// TIA Portal V20 export
FUNCTION_BLOCK "PR_TT-1MasterSeq_Soft2.0_workflow_b380e4"   // FB53, LAD
{ S7_Optimized_Access := 'TRUE' }
// stored: MemoryReserve 100, SetENOAutomatically false
   VAR_INPUT
      iAllStationProcessOver : Bool;
      iAutoRunning : Bool;
      iHiPotTestOver_1 : Bool;
      iHiPotTestOver_2 : Bool;
      iHiPot_RTR_1 : Bool;
      iHiPot_RTR_2 : Bool;
      iIndexOver : Bool;
      iIndex_RTR_Place1 : Bool;
      iIndex_RTR_Place2 : Bool;
      iOTS_Frm_Shuttle_1 : Bool;
      iOTS_Frm_Shuttle_2 : Bool;
      iOTS_Frm_TransferGantry : Bool;
      iOperatorAck : Bool;
      iPartPickOver : Bool;
      iPartPickOver_1 : Bool;
      iPartPickOver_2 : Bool;
      iPartPlaceByTransferGantry : Bool;
      iPartPlaceOver_IFGantry : Bool;
      iPartPlaceOver_IndexPlace1 : Bool;
      iPartPlaceOver_IndexPlace2 : Bool;
      iPartPresent_IFGantry : Bool;
      iPartPresent_Shuttle_1 : Bool;
      iPartPresent_Shuttle_2 : Bool;
      iPartPresent_TxGantry_1 : Bool;
      iPartPresent_TxGantry_2 : Bool;
      iRTR_Frm_TransferGantry_1 : Bool;
      iRTR_Frm_TransferGantry_2 : Bool;
      iReset_fault : Bool;
      iShuttleReadyToReceive : Bool;
      iSstMode : Bool;
      iSstPB : Bool;
   END_VAR
   VAR_OUTPUT
      qError : Array[1..1] of Bool;
      qInfeedGantry_PickStart : Bool;
      qInfeedGantry_PlaceStart : Bool;
      qShuttle_1PickStart : Bool;
      qShuttle_1PlaceStart : Bool;
      qShuttle_2PickStart : Bool;
      qShuttle_2PlaceStart : Bool;
      qTransferGantry1_PickStart : Bool;
      qTransferGantry1_PlaceStart : Bool;
      qTransferGantry2_PickStart : Bool;
      qTransferGantry2_PlaceStart : Bool;
   END_VAR
   VAR
      c10_ChkPartStsAtSubStn_T1 : Bool;
      c10_ChkPartStsAtSubStn_T2 : Bool;
      c10_ChkPartStsAtSubStn_T3 : Bool;
      c10_ChkPartStsAtSubStn_T4 : Bool;
      c10_ChkPartStsAtSubStn_T5 : Bool;
      c10_ChkPartStsAtSubStn_T6 : Bool;
      c10_ChkPartStsAtSubStn_T7 : Bool;
      c130_ChkPartPrsntStsShuttle2_T1 : Bool;
      c130_ChkPartPrsntStsShuttle2_T2 : Bool;
      c200_ChkPartPrsntTxGantry1_T1 : Bool;
      c200_ChkPartPrsntTxGantry1_T2 : Bool;
      c250_ChkPartPrsntTxGantry2_T1 : Bool;
      c250_ChkPartPrsntTxGantry2_T2 : Bool;
      c300_ChkPartPrsntIndexer_T1 : Bool;
      c300_ChkPartPrsntIndexer_T2 : Bool;
      c30_ChkPartStsIFGantry_T1 : Bool;
      c30_ChkPartStsIFGantry_T2 : Bool;
      c70_ChkPartPrsntStsShuttle1_T1 : Bool;
      c70_ChkPartPrsntStsShuttle1_T2 : Bool;
      StateNo : Int;
      s100_WtHiPotTestOver1 : Bool;
      s100_WtHiPotTestOver1_T1 : Bool;
      s10_ChkPartStsAtSubStn : Bool;
      s10_ChkPartStsAtSubStn_T1 : Bool;
      s10_ChkPartStsAtSubStn_T2 : Bool;
      s10_ChkPartStsAtSubStn_T3 : Bool;
      s10_ChkPartStsAtSubStn_T4 : Bool;
      s10_ChkPartStsAtSubStn_T5 : Bool;
      s10_ChkPartStsAtSubStn_T6 : Bool;
      s10_ChkPartStsAtSubStn_T7 : Bool;
      s110_WtTxGantryRTR1 : Bool;
      s110_WtTxGantryRTR1_T1 : Bool;
      s120_WtPartUnldOvrTxGantry1 : Bool;
      s120_WtPartUnldOvrTxGantry1_T1 : Bool;
      s130_ChkPartPrsntStsShuttle2 : Bool;
      s130_ChkPartPrsntStsShuttle2_T1 : Bool;
      s130_ChkPartPrsntStsShuttle2_T2 : Bool;
      s140_WtIFGantryPlacePart2 : Bool;
      s140_WtIFGantryPlacePart2_T1 : Bool;
      s150_WtHiPotRdyRcvPart2 : Bool;
      s150_WtHiPotRdyRcvPart2_T1 : Bool;
      s160_WtHiPotTestOver2 : Bool;
      s160_WtHiPotTestOver2_T1 : Bool;
      s170_WtTxGantryRTR2 : Bool;
      s170_WtTxGantryRTR2_T1 : Bool;
      s190_WtPartUnldOvrTxGantry2 : Bool;
      s190_WtPartUnldOvrTxGantry2_T1 : Bool;
      s1_WtResetRel : Bool;
      s1_WtResetRel_T1 : Bool;
      s200_ChkPartPrsntTxGantry1 : Bool;
      s200_ChkPartPrsntTxGantry1_T1 : Bool;
      s200_ChkPartPrsntTxGantry1_T2 : Bool;
      s20_WtOperatorAck : Bool;
      s20_WtOperatorAck_T1 : Bool;
      s210_WtShuttle1RdySendPal : Bool;
      s210_WtShuttle1RdySendPal_T1 : Bool;
      s220_WtPartPickTxGantry1 : Bool;
      s220_WtPartPickTxGantry1_T1 : Bool;
      s230_WtIndexRTRPlace1 : Bool;
      s230_WtIndexRTRPlace1_T1 : Bool;
      s240_WtPartPlaceOverIndexPlace1 : Bool;
      s240_WtPartPlaceOverIndexPlace1_T1 : Bool;
      s250_ChkPartPrsntTxGantry2 : Bool;
      s250_ChkPartPrsntTxGantry2_T1 : Bool;
      s250_ChkPartPrsntTxGantry2_T2 : Bool;
      s260_WtShuttle2RdySendPal : Bool;
      s260_WtShuttle2RdySendPal_T1 : Bool;
      s270_WtPartPickTxGantry2 : Bool;
      s270_WtPartPickTxGantry2_T1 : Bool;
      s280_WtIndexRTRPlace2 : Bool;
      s280_WtIndexRTRPlace2_T1 : Bool;
      s290_WtPartPlaceOverIndexPlace2 : Bool;
      s290_WtPartPlaceOverIndexPlace2_T1 : Bool;
      s300_ChkPartPrsntIndexer : Bool;
      s300_ChkPartPrsntIndexer_T1 : Bool;
      s300_ChkPartPrsntIndexer_T2 : Bool;
      s30_ChkPartStsIFGantry : Bool;
      s30_ChkPartStsIFGantry_T1 : Bool;
      s30_ChkPartStsIFGantry_T2 : Bool;
      s310_WtOTSFrmTxGantry : Bool;
      s310_WtOTSFrmTxGantry_T1 : Bool;
      s320_WtPartPlaceByTxGantry : Bool;
      s320_WtPartPlaceByTxGantry_T1 : Bool;
      s330_WtAllStnProcessOver : Bool;
      s330_WtAllStnProcessOver_T1 : Bool;
      s340_WtIndexOver : Bool;
      s340_WtIndexOver_T1 : Bool;
      s40_WtPartPickOverIFGantry : Bool;
      s40_WtPartPickOverIFGantry_T1 : Bool;
      s50_WtShuttleRdyRcvPart : Bool;
      s50_WtShuttleRdyRcvPart_T1 : Bool;
      s60_WtPartPlaceByGantry : Bool;
      s60_WtPartPlaceByGantry_T1 : Bool;
      s70_ChkPartPrsntStsShuttle1 : Bool;
      s70_ChkPartPrsntStsShuttle1_T1 : Bool;
      s70_ChkPartPrsntStsShuttle1_T2 : Bool;
      s80_WtIFGantryPlacePart : Bool;
      s80_WtIFGantryPlacePart_T1 : Bool;
      s90_WtHiPotRdyRcvPart1 : Bool;
      s90_WtHiPotRdyRcvPart1_T1 : Bool;
      sAbnormalCondition : Bool;
      sIndexerSeq : Bool;
      sInfeedGantry : Bool;
      sPartAbsentAtAllStn : Bool;
      sPartPrsntAtStn : Bool;
      sShuttle_1Seq : Bool;
      sShuttle_2Seq : Bool;
      sSst : Bool;
      sSstPulse : Bool;
      sSstRise : Bool;
      sStWtResetRel : Bool;
      sStWtResetRel_T1 : Bool;
      sTransferGantry_1Seq : Bool;
      sTransferGantry_2Seq : Bool;
   END_VAR
   VAR_TEMP
      tOne : Bool;
   END_VAR
   VAR_TEMP   // added for the SCL form of the ladder/FBD networks
      _w1 : Bool;
      _w2 : Bool;
      _w3 : Bool;
      _w4 : Bool;
      _w5 : Bool;
      _w6 : Bool;
   END_VAR
BEGIN

REGION Network 1
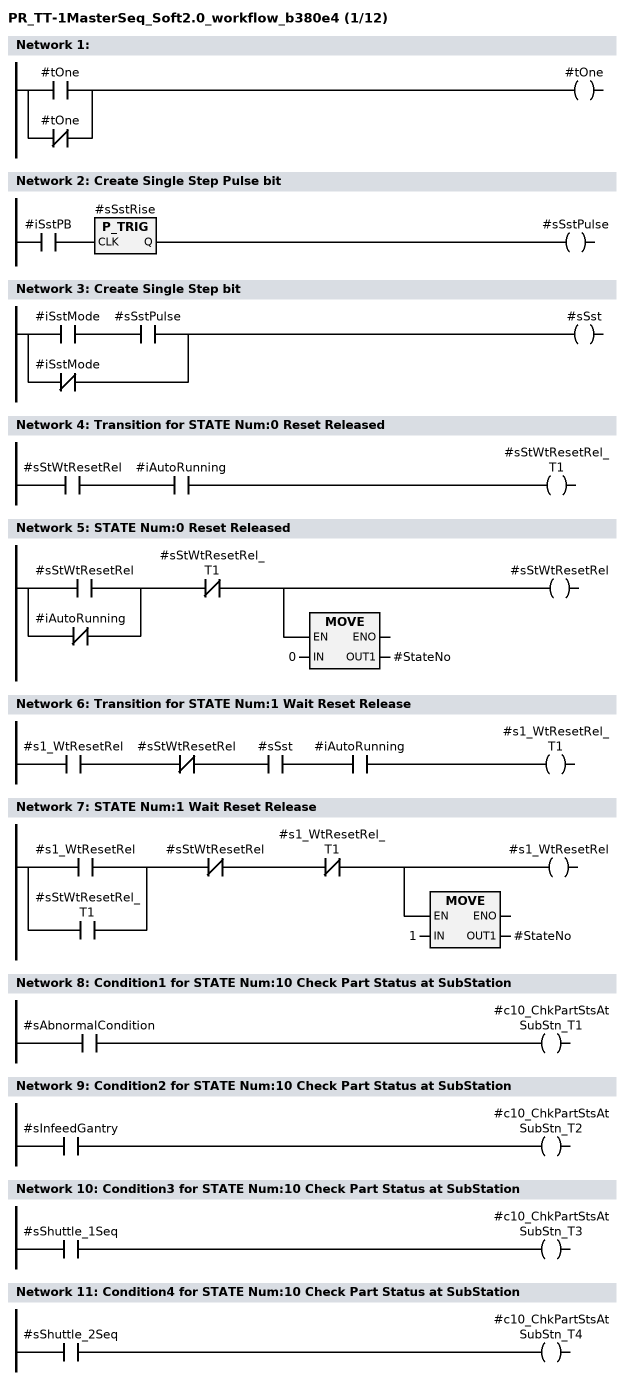
   RUNG wire#powerrail
      Contact( #tOne )
      wire#w1
      Coil( #tOne )
   END_RUNG
   RUNG wire#powerrail
      I_Contact( #tOne )
   END_RUNG wire#w1
   // the same network as SCL:
   #tOne := #tOne OR NOT #tOne;
END_REGION

REGION Network 2: Create Single Step Pulse bit
   RUNG wire#powerrail
      Contact( #iSstPB )
      P_Trig( #sSstRise )
      Coil( #sSstPulse )
   END_RUNG
   // the same network as SCL:
   #_w1 := #iSstPB AND NOT #sSstRise;   // rising edge
   #sSstRise := #iSstPB;
   #sSstPulse := #_w1;
END_REGION

REGION Network 3: Create Single Step bit
   RUNG wire#powerrail
      Contact( #iSstMode )
      Contact( #sSstPulse )
      wire#w1
      Coil( #sSst )
   END_RUNG
   RUNG wire#powerrail
      I_Contact( #iSstMode )
   END_RUNG wire#w1
   // the same network as SCL:
   #sSst := (#iSstMode AND #sSstPulse) OR NOT #iSstMode;
END_REGION

REGION Network 4: Transition for STATE Num:0 Reset Released
   RUNG wire#powerrail
      Contact( #sStWtResetRel )
      Contact( #iAutoRunning )
      Coil( #sStWtResetRel_T1 )
   END_RUNG
   // the same network as SCL:
   #sStWtResetRel_T1 := #sStWtResetRel AND #iAutoRunning;
END_REGION

REGION Network 5: STATE Num:0 Reset Released
   RUNG wire#powerrail
      Contact( #sStWtResetRel )
      wire#w1
      I_Contact( #sStWtResetRel_T1 )
      wire#w2
      Coil( #sStWtResetRel )
   END_RUNG
   RUNG wire#powerrail
      I_Contact( #iAutoRunning )
   END_RUNG wire#w1
   RUNG wire#w2
      { S7_GenerateENO := "TRUE" } Move(in := 0, out1 => #StateNo)
   END_RUNG
   // the same network as SCL:
   #sStWtResetRel := (#sStWtResetRel OR NOT #iAutoRunning) AND NOT #sStWtResetRel_T1;
   IF #sStWtResetRel THEN #StateNo := 0; END_IF;
END_REGION

REGION Network 6: Transition for STATE Num:1 Wait Reset Release
   RUNG wire#powerrail
      Contact( #s1_WtResetRel )
      I_Contact( #sStWtResetRel )
      Contact( #sSst )
      Contact( #iAutoRunning )
      Coil( #s1_WtResetRel_T1 )
   END_RUNG
   // the same network as SCL:
   #s1_WtResetRel_T1 := #s1_WtResetRel AND NOT #sStWtResetRel AND #sSst AND #iAutoRunning;
END_REGION

REGION Network 7: STATE Num:1 Wait Reset Release
   RUNG wire#powerrail
      Contact( #s1_WtResetRel )
      wire#w1
      I_Contact( #sStWtResetRel )
      I_Contact( #s1_WtResetRel_T1 )
      wire#w2
      Coil( #s1_WtResetRel )
   END_RUNG
   RUNG wire#powerrail
      Contact( #sStWtResetRel_T1 )
   END_RUNG wire#w1
   RUNG wire#w2
      { S7_GenerateENO := "TRUE" } Move(in := 1, out1 => #StateNo)
   END_RUNG
   // the same network as SCL:
   #s1_WtResetRel := (#s1_WtResetRel OR #sStWtResetRel_T1) AND NOT #sStWtResetRel AND NOT #s1_WtResetRel_T1;
   IF #s1_WtResetRel THEN #StateNo := 1; END_IF;
END_REGION

REGION Network 8: Condition1 for STATE Num:10 Check Part Status at SubStation
   RUNG wire#powerrail
      Contact( #sAbnormalCondition )
      Coil( #c10_ChkPartStsAtSubStn_T1 )
   END_RUNG
   // the same network as SCL:
   #c10_ChkPartStsAtSubStn_T1 := #sAbnormalCondition;
END_REGION

REGION Network 9: Condition2 for STATE Num:10 Check Part Status at SubStation
   RUNG wire#powerrail
      Contact( #sInfeedGantry )
      Coil( #c10_ChkPartStsAtSubStn_T2 )
   END_RUNG
   // the same network as SCL:
   #c10_ChkPartStsAtSubStn_T2 := #sInfeedGantry;
END_REGION

REGION Network 10: Condition3 for STATE Num:10 Check Part Status at SubStation
   RUNG wire#powerrail
      Contact( #sShuttle_1Seq )
      Coil( #c10_ChkPartStsAtSubStn_T3 )
   END_RUNG
   // the same network as SCL:
   #c10_ChkPartStsAtSubStn_T3 := #sShuttle_1Seq;
END_REGION

REGION Network 11: Condition4 for STATE Num:10 Check Part Status at SubStation
   RUNG wire#powerrail
      Contact( #sShuttle_2Seq )
      Coil( #c10_ChkPartStsAtSubStn_T4 )
   END_RUNG
   // the same network as SCL:
   #c10_ChkPartStsAtSubStn_T4 := #sShuttle_2Seq;
END_REGION

REGION Network 12: Condition5 for STATE Num:10 Check Part Status at SubStation
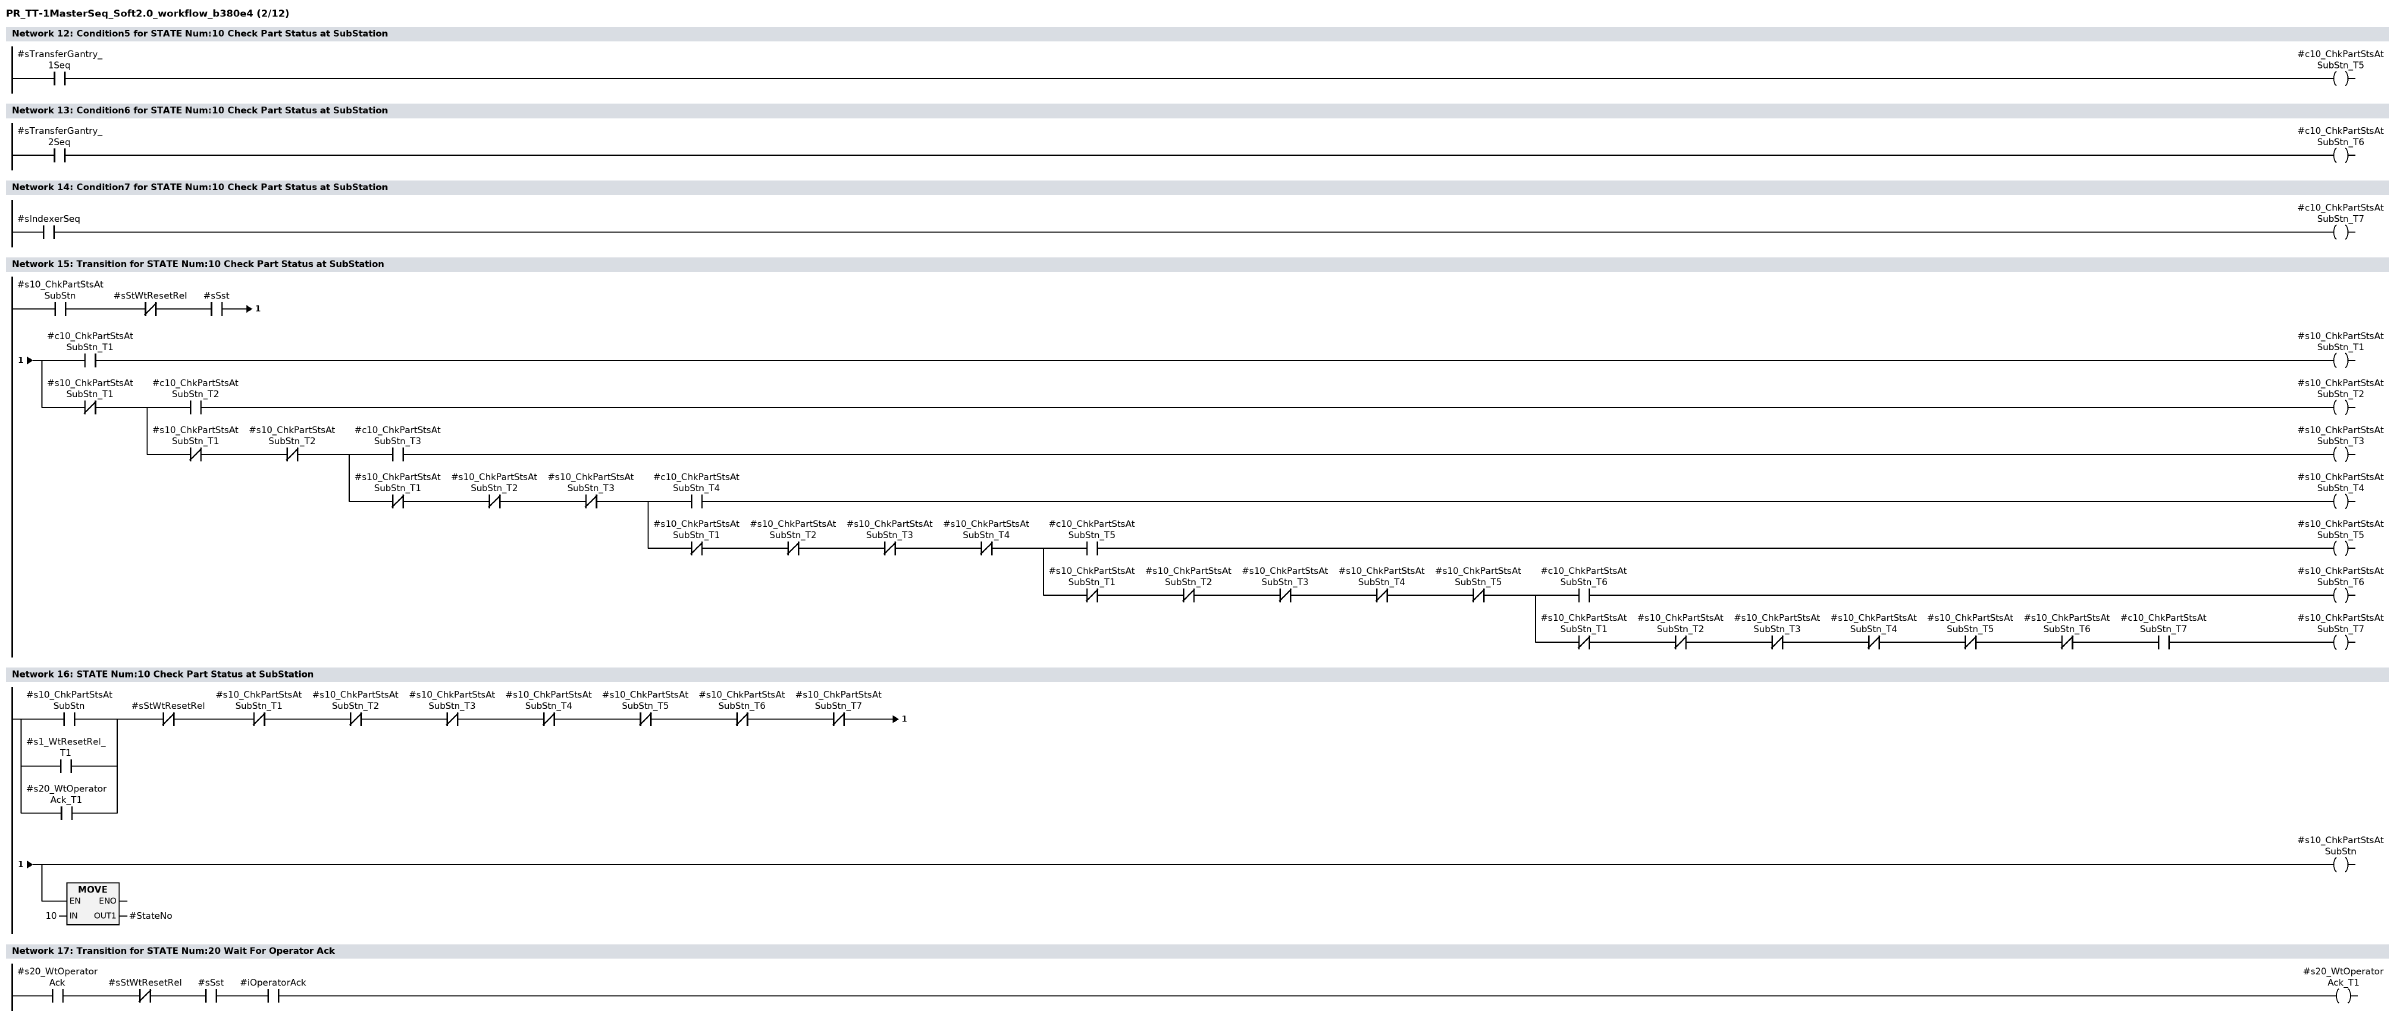
   RUNG wire#powerrail
      Contact( #sTransferGantry_1Seq )
      Coil( #c10_ChkPartStsAtSubStn_T5 )
   END_RUNG
   // the same network as SCL:
   #c10_ChkPartStsAtSubStn_T5 := #sTransferGantry_1Seq;
END_REGION

REGION Network 13: Condition6 for STATE Num:10 Check Part Status at SubStation
   RUNG wire#powerrail
      Contact( #sTransferGantry_2Seq )
      Coil( #c10_ChkPartStsAtSubStn_T6 )
   END_RUNG
   // the same network as SCL:
   #c10_ChkPartStsAtSubStn_T6 := #sTransferGantry_2Seq;
END_REGION

REGION Network 14: Condition7 for STATE Num:10 Check Part Status at SubStation
   RUNG wire#powerrail
      Contact( #sIndexerSeq )
      Coil( #c10_ChkPartStsAtSubStn_T7 )
   END_RUNG
   // the same network as SCL:
   #c10_ChkPartStsAtSubStn_T7 := #sIndexerSeq;
END_REGION

REGION Network 15: Transition for STATE Num:10 Check Part Status at SubStation
   RUNG wire#powerrail
      Contact( #s10_ChkPartStsAtSubStn )
      I_Contact( #sStWtResetRel )
      Contact( #sSst )
      wire#w1
      Contact( #c10_ChkPartStsAtSubStn_T1 )
      Coil( #s10_ChkPartStsAtSubStn_T1 )
   END_RUNG
   RUNG wire#w1
      I_Contact( #s10_ChkPartStsAtSubStn_T1 )
      wire#w2
      Contact( #c10_ChkPartStsAtSubStn_T2 )
      Coil( #s10_ChkPartStsAtSubStn_T2 )
   END_RUNG
   RUNG wire#w2
      I_Contact( #s10_ChkPartStsAtSubStn_T1 )
      I_Contact( #s10_ChkPartStsAtSubStn_T2 )
      wire#w3
      Contact( #c10_ChkPartStsAtSubStn_T3 )
      Coil( #s10_ChkPartStsAtSubStn_T3 )
   END_RUNG
   RUNG wire#w3
      I_Contact( #s10_ChkPartStsAtSubStn_T1 )
      I_Contact( #s10_ChkPartStsAtSubStn_T2 )
      I_Contact( #s10_ChkPartStsAtSubStn_T3 )
      wire#w4
      Contact( #c10_ChkPartStsAtSubStn_T4 )
      Coil( #s10_ChkPartStsAtSubStn_T4 )
   END_RUNG
   RUNG wire#w4
      I_Contact( #s10_ChkPartStsAtSubStn_T1 )
      I_Contact( #s10_ChkPartStsAtSubStn_T2 )
      I_Contact( #s10_ChkPartStsAtSubStn_T3 )
      I_Contact( #s10_ChkPartStsAtSubStn_T4 )
      wire#w5
      Contact( #c10_ChkPartStsAtSubStn_T5 )
      Coil( #s10_ChkPartStsAtSubStn_T5 )
   END_RUNG
   RUNG wire#w5
      I_Contact( #s10_ChkPartStsAtSubStn_T1 )
      I_Contact( #s10_ChkPartStsAtSubStn_T2 )
      I_Contact( #s10_ChkPartStsAtSubStn_T3 )
      I_Contact( #s10_ChkPartStsAtSubStn_T4 )
      I_Contact( #s10_ChkPartStsAtSubStn_T5 )
      wire#w6
      Contact( #c10_ChkPartStsAtSubStn_T6 )
      Coil( #s10_ChkPartStsAtSubStn_T6 )
   END_RUNG
   RUNG wire#w6
      I_Contact( #s10_ChkPartStsAtSubStn_T1 )
      I_Contact( #s10_ChkPartStsAtSubStn_T2 )
      I_Contact( #s10_ChkPartStsAtSubStn_T3 )
      I_Contact( #s10_ChkPartStsAtSubStn_T4 )
      I_Contact( #s10_ChkPartStsAtSubStn_T5 )
      I_Contact( #s10_ChkPartStsAtSubStn_T6 )
      Contact( #c10_ChkPartStsAtSubStn_T7 )
      Coil( #s10_ChkPartStsAtSubStn_T7 )
   END_RUNG
   // the same network as SCL:
   #_w1 := #s10_ChkPartStsAtSubStn AND NOT #sStWtResetRel AND #sSst;
   #s10_ChkPartStsAtSubStn_T1 := #_w1 AND #c10_ChkPartStsAtSubStn_T1;
   #_w2 := #_w1 AND NOT #s10_ChkPartStsAtSubStn_T1;
   #s10_ChkPartStsAtSubStn_T2 := #_w2 AND #c10_ChkPartStsAtSubStn_T2;
   #_w3 := #_w2 AND NOT #s10_ChkPartStsAtSubStn_T1 AND NOT #s10_ChkPartStsAtSubStn_T2;
   #s10_ChkPartStsAtSubStn_T3 := #_w3 AND #c10_ChkPartStsAtSubStn_T3;
   #_w4 := #_w3 AND NOT #s10_ChkPartStsAtSubStn_T1 AND NOT #s10_ChkPartStsAtSubStn_T2 AND NOT #s10_ChkPartStsAtSubStn_T3;
   #s10_ChkPartStsAtSubStn_T4 := #_w4 AND #c10_ChkPartStsAtSubStn_T4;
   #_w5 := #_w4 AND NOT #s10_ChkPartStsAtSubStn_T1 AND NOT #s10_ChkPartStsAtSubStn_T2 AND NOT #s10_ChkPartStsAtSubStn_T3 AND NOT #s10_ChkPartStsAtSubStn_T4;
   #s10_ChkPartStsAtSubStn_T5 := #_w5 AND #c10_ChkPartStsAtSubStn_T5;
   #_w6 := #_w5 AND NOT #s10_ChkPartStsAtSubStn_T1 AND NOT #s10_ChkPartStsAtSubStn_T2 AND NOT #s10_ChkPartStsAtSubStn_T3 AND NOT #s10_ChkPartStsAtSubStn_T4 AND NOT #s10_ChkPartStsAtSubStn_T5;
   #s10_ChkPartStsAtSubStn_T6 := #_w6 AND #c10_ChkPartStsAtSubStn_T6;
   #s10_ChkPartStsAtSubStn_T7 := #_w6 AND NOT #s10_ChkPartStsAtSubStn_T1 AND NOT #s10_ChkPartStsAtSubStn_T2 AND NOT #s10_ChkPartStsAtSubStn_T3 AND NOT #s10_ChkPartStsAtSubStn_T4 AND NOT #s10_ChkPartStsAtSubStn_T5 AND NOT #s10_ChkPartStsAtSubStn_T6 AND #c10_ChkPartStsAtSubStn_T7;
END_REGION

REGION Network 16: STATE Num:10 Check Part Status at SubStation
   RUNG wire#powerrail
      Contact( #s10_ChkPartStsAtSubStn )
      wire#w1
      I_Contact( #sStWtResetRel )
      I_Contact( #s10_ChkPartStsAtSubStn_T1 )
      I_Contact( #s10_ChkPartStsAtSubStn_T2 )
      I_Contact( #s10_ChkPartStsAtSubStn_T3 )
      I_Contact( #s10_ChkPartStsAtSubStn_T4 )
      I_Contact( #s10_ChkPartStsAtSubStn_T5 )
      I_Contact( #s10_ChkPartStsAtSubStn_T6 )
      I_Contact( #s10_ChkPartStsAtSubStn_T7 )
      wire#w2
      Coil( #s10_ChkPartStsAtSubStn )
   END_RUNG
   RUNG wire#powerrail
      Contact( #s1_WtResetRel_T1 )
   END_RUNG wire#w1
   RUNG wire#powerrail
      Contact( #s20_WtOperatorAck_T1 )
   END_RUNG wire#w1
   RUNG wire#w2
      { S7_GenerateENO := "TRUE" } Move(in := 10, out1 => #StateNo)
   END_RUNG
   // the same network as SCL:
   #s10_ChkPartStsAtSubStn := (#s10_ChkPartStsAtSubStn OR #s1_WtResetRel_T1 OR #s20_WtOperatorAck_T1) AND NOT #sStWtResetRel AND NOT #s10_ChkPartStsAtSubStn_T1 AND NOT #s10_ChkPartStsAtSubStn_T2 AND NOT #s10_ChkPartStsAtSubStn_T3 AND NOT #s10_ChkPartStsAtSubStn_T4 AND NOT #s10_ChkPartStsAtSubStn_T5 AND NOT #s10_ChkPartStsAtSubStn_T6 AND NOT #s10_ChkPartStsAtSubStn_T7;
   IF #s10_ChkPartStsAtSubStn THEN #StateNo := 10; END_IF;
END_REGION

REGION Network 17: Transition for STATE Num:20 Wait For Operator Ack
   RUNG wire#powerrail
      Contact( #s20_WtOperatorAck )
      I_Contact( #sStWtResetRel )
      Contact( #sSst )
      Contact( #iOperatorAck )
      Coil( #s20_WtOperatorAck_T1 )
   END_RUNG
   // the same network as SCL:
   #s20_WtOperatorAck_T1 := #s20_WtOperatorAck AND NOT #sStWtResetRel AND #sSst AND #iOperatorAck;
END_REGION

REGION Network 18: STATE Num:20 Wait For Operator Ack
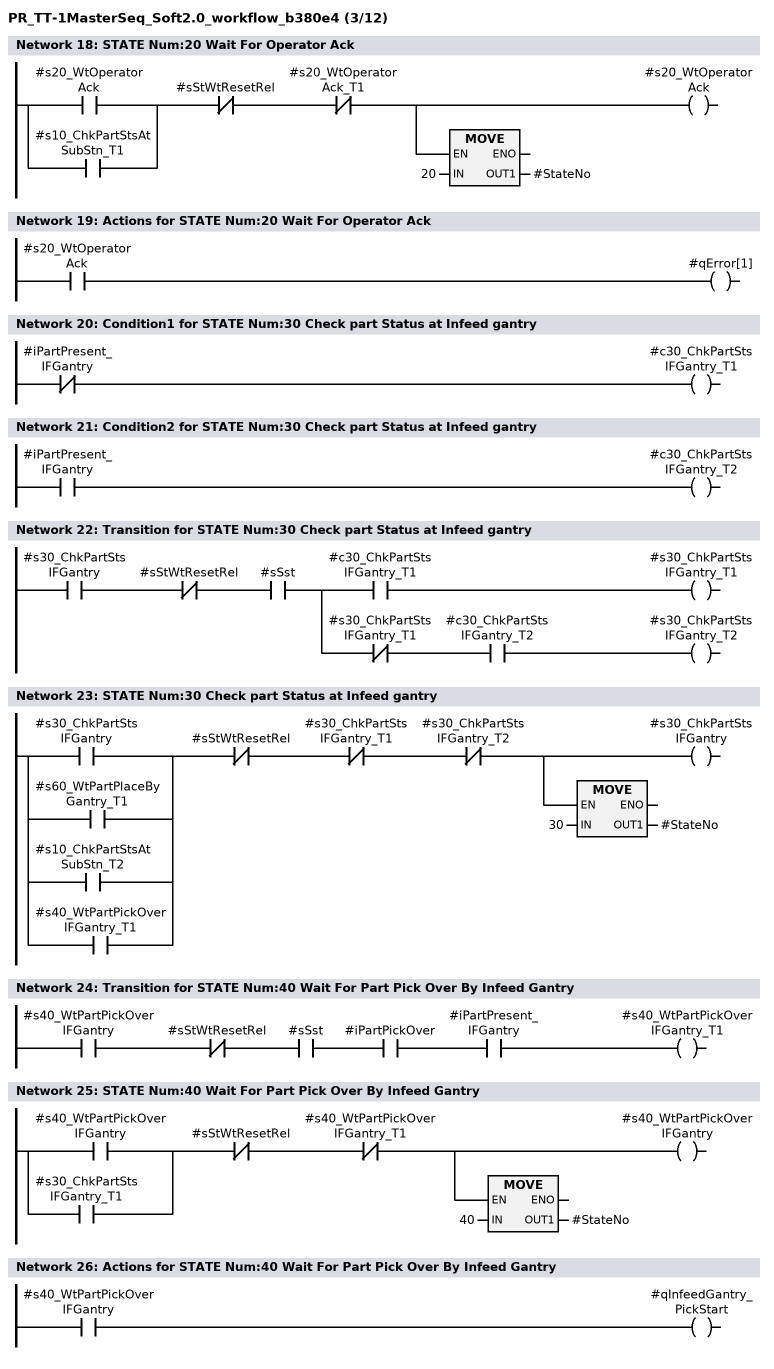
   RUNG wire#powerrail
      Contact( #s20_WtOperatorAck )
      wire#w1
      I_Contact( #sStWtResetRel )
      I_Contact( #s20_WtOperatorAck_T1 )
      wire#w2
      Coil( #s20_WtOperatorAck )
   END_RUNG
   RUNG wire#powerrail
      Contact( #s10_ChkPartStsAtSubStn_T1 )
   END_RUNG wire#w1
   RUNG wire#w2
      { S7_GenerateENO := "TRUE" } Move(in := 20, out1 => #StateNo)
   END_RUNG
   // the same network as SCL:
   #s20_WtOperatorAck := (#s20_WtOperatorAck OR #s10_ChkPartStsAtSubStn_T1) AND NOT #sStWtResetRel AND NOT #s20_WtOperatorAck_T1;
   IF #s20_WtOperatorAck THEN #StateNo := 20; END_IF;
END_REGION

REGION Network 19: Actions for STATE Num:20 Wait For Operator Ack
   RUNG wire#powerrail
      Contact( #s20_WtOperatorAck )
      Coil( #qError[1] )
   END_RUNG
   // the same network as SCL:
   #qError[1] := #s20_WtOperatorAck;
END_REGION

REGION Network 20: Condition1 for STATE Num:30 Check part Status at Infeed gantry
   RUNG wire#powerrail
      I_Contact( #iPartPresent_IFGantry )
      Coil( #c30_ChkPartStsIFGantry_T1 )
   END_RUNG
   // the same network as SCL:
   #c30_ChkPartStsIFGantry_T1 := NOT #iPartPresent_IFGantry;
END_REGION

REGION Network 21: Condition2 for STATE Num:30 Check part Status at Infeed gantry
   RUNG wire#powerrail
      Contact( #iPartPresent_IFGantry )
      Coil( #c30_ChkPartStsIFGantry_T2 )
   END_RUNG
   // the same network as SCL:
   #c30_ChkPartStsIFGantry_T2 := #iPartPresent_IFGantry;
END_REGION

REGION Network 22: Transition for STATE Num:30 Check part Status at Infeed gantry
   RUNG wire#powerrail
      Contact( #s30_ChkPartStsIFGantry )
      I_Contact( #sStWtResetRel )
      Contact( #sSst )
      wire#w1
      Contact( #c30_ChkPartStsIFGantry_T1 )
      Coil( #s30_ChkPartStsIFGantry_T1 )
   END_RUNG
   RUNG wire#w1
      I_Contact( #s30_ChkPartStsIFGantry_T1 )
      Contact( #c30_ChkPartStsIFGantry_T2 )
      Coil( #s30_ChkPartStsIFGantry_T2 )
   END_RUNG
   // the same network as SCL:
   #_w1 := #s30_ChkPartStsIFGantry AND NOT #sStWtResetRel AND #sSst;
   #s30_ChkPartStsIFGantry_T1 := #_w1 AND #c30_ChkPartStsIFGantry_T1;
   #s30_ChkPartStsIFGantry_T2 := #_w1 AND NOT #s30_ChkPartStsIFGantry_T1 AND #c30_ChkPartStsIFGantry_T2;
END_REGION

REGION Network 23: STATE Num:30 Check part Status at Infeed gantry
   RUNG wire#powerrail
      Contact( #s30_ChkPartStsIFGantry )
      wire#w1
      I_Contact( #sStWtResetRel )
      I_Contact( #s30_ChkPartStsIFGantry_T1 )
      I_Contact( #s30_ChkPartStsIFGantry_T2 )
      wire#w2
      Coil( #s30_ChkPartStsIFGantry )
   END_RUNG
   RUNG wire#powerrail
      Contact( #s60_WtPartPlaceByGantry_T1 )
   END_RUNG wire#w1
   RUNG wire#powerrail
      Contact( #s10_ChkPartStsAtSubStn_T2 )
   END_RUNG wire#w1
   RUNG wire#powerrail
      Contact( #s40_WtPartPickOverIFGantry_T1 )
   END_RUNG wire#w1
   RUNG wire#w2
      { S7_GenerateENO := "TRUE" } Move(in := 30, out1 => #StateNo)
   END_RUNG
   // the same network as SCL:
   #s30_ChkPartStsIFGantry := (#s30_ChkPartStsIFGantry OR #s60_WtPartPlaceByGantry_T1 OR #s10_ChkPartStsAtSubStn_T2 OR #s40_WtPartPickOverIFGantry_T1) AND NOT #sStWtResetRel AND NOT #s30_ChkPartStsIFGantry_T1 AND NOT #s30_ChkPartStsIFGantry_T2;
   IF #s30_ChkPartStsIFGantry THEN #StateNo := 30; END_IF;
END_REGION

REGION Network 24: Transition for STATE Num:40 Wait For Part Pick Over By Infeed Gantry
   RUNG wire#powerrail
      Contact( #s40_WtPartPickOverIFGantry )
      I_Contact( #sStWtResetRel )
      Contact( #sSst )
      Contact( #iPartPickOver )
      Contact( #iPartPresent_IFGantry )
      Coil( #s40_WtPartPickOverIFGantry_T1 )
   END_RUNG
   // the same network as SCL:
   #s40_WtPartPickOverIFGantry_T1 := #s40_WtPartPickOverIFGantry AND NOT #sStWtResetRel AND #sSst AND #iPartPickOver AND #iPartPresent_IFGantry;
END_REGION

REGION Network 25: STATE Num:40 Wait For Part Pick Over By Infeed Gantry
   RUNG wire#powerrail
      Contact( #s40_WtPartPickOverIFGantry )
      wire#w1
      I_Contact( #sStWtResetRel )
      I_Contact( #s40_WtPartPickOverIFGantry_T1 )
      wire#w2
      Coil( #s40_WtPartPickOverIFGantry )
   END_RUNG
   RUNG wire#powerrail
      Contact( #s30_ChkPartStsIFGantry_T1 )
   END_RUNG wire#w1
   RUNG wire#w2
      { S7_GenerateENO := "TRUE" } Move(in := 40, out1 => #StateNo)
   END_RUNG
   // the same network as SCL:
   #s40_WtPartPickOverIFGantry := (#s40_WtPartPickOverIFGantry OR #s30_ChkPartStsIFGantry_T1) AND NOT #sStWtResetRel AND NOT #s40_WtPartPickOverIFGantry_T1;
   IF #s40_WtPartPickOverIFGantry THEN #StateNo := 40; END_IF;
END_REGION

REGION Network 26: Actions for STATE Num:40 Wait For Part Pick Over By Infeed Gantry
   RUNG wire#powerrail
      Contact( #s40_WtPartPickOverIFGantry )
      Coil( #qInfeedGantry_PickStart )
   END_RUNG
   // the same network as SCL:
   #qInfeedGantry_PickStart := #s40_WtPartPickOverIFGantry;
END_REGION

REGION Network 27: Transition for STATE Num:50 Wait Shuttle Ready To Receive Part
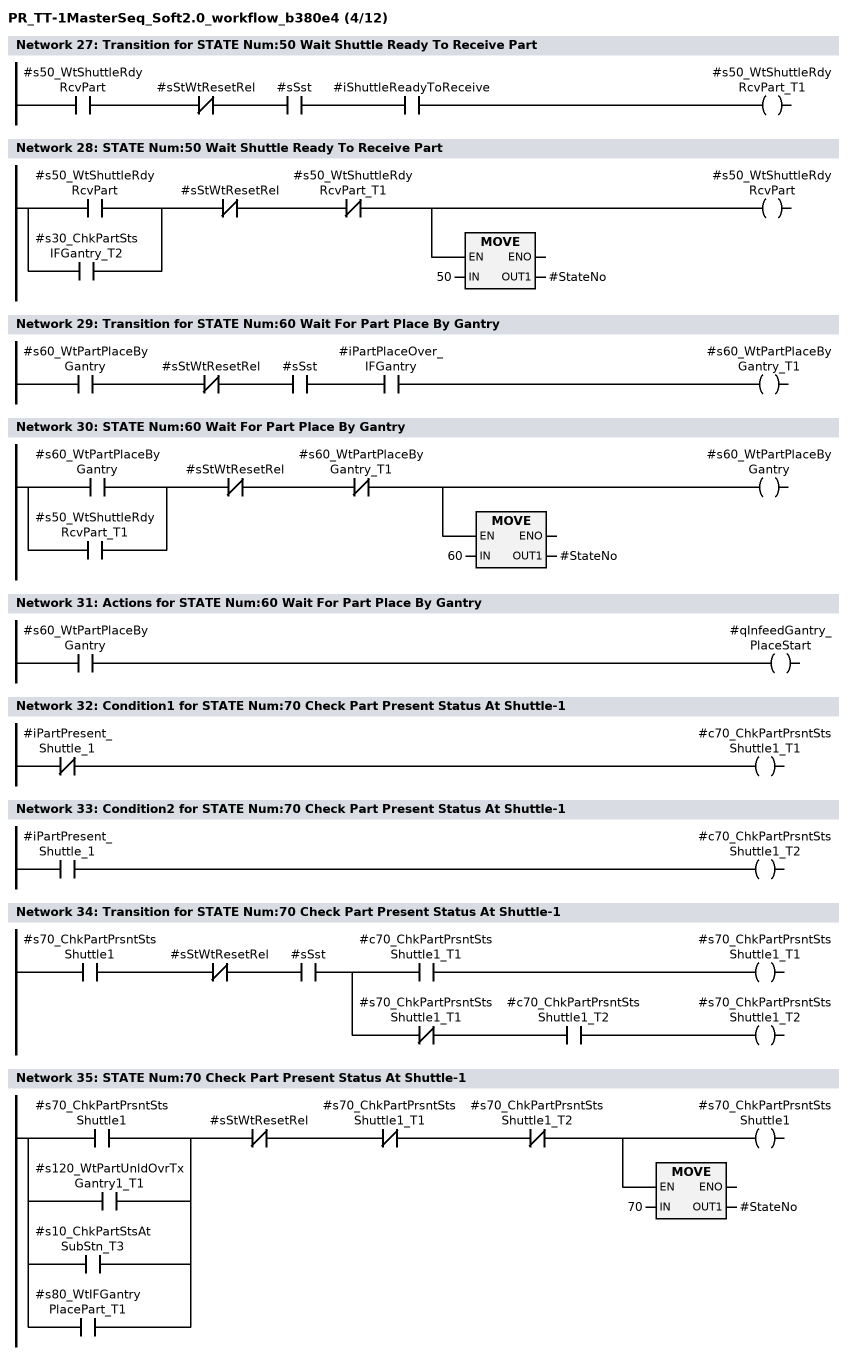
   RUNG wire#powerrail
      Contact( #s50_WtShuttleRdyRcvPart )
      I_Contact( #sStWtResetRel )
      Contact( #sSst )
      Contact( #iShuttleReadyToReceive )
      Coil( #s50_WtShuttleRdyRcvPart_T1 )
   END_RUNG
   // the same network as SCL:
   #s50_WtShuttleRdyRcvPart_T1 := #s50_WtShuttleRdyRcvPart AND NOT #sStWtResetRel AND #sSst AND #iShuttleReadyToReceive;
END_REGION

REGION Network 28: STATE Num:50 Wait Shuttle Ready To Receive Part
   RUNG wire#powerrail
      Contact( #s50_WtShuttleRdyRcvPart )
      wire#w1
      I_Contact( #sStWtResetRel )
      I_Contact( #s50_WtShuttleRdyRcvPart_T1 )
      wire#w2
      Coil( #s50_WtShuttleRdyRcvPart )
   END_RUNG
   RUNG wire#powerrail
      Contact( #s30_ChkPartStsIFGantry_T2 )
   END_RUNG wire#w1
   RUNG wire#w2
      { S7_GenerateENO := "TRUE" } Move(in := 50, out1 => #StateNo)
   END_RUNG
   // the same network as SCL:
   #s50_WtShuttleRdyRcvPart := (#s50_WtShuttleRdyRcvPart OR #s30_ChkPartStsIFGantry_T2) AND NOT #sStWtResetRel AND NOT #s50_WtShuttleRdyRcvPart_T1;
   IF #s50_WtShuttleRdyRcvPart THEN #StateNo := 50; END_IF;
END_REGION

REGION Network 29: Transition for STATE Num:60 Wait For Part Place By Gantry
   RUNG wire#powerrail
      Contact( #s60_WtPartPlaceByGantry )
      I_Contact( #sStWtResetRel )
      Contact( #sSst )
      Contact( #iPartPlaceOver_IFGantry )
      Coil( #s60_WtPartPlaceByGantry_T1 )
   END_RUNG
   // the same network as SCL:
   #s60_WtPartPlaceByGantry_T1 := #s60_WtPartPlaceByGantry AND NOT #sStWtResetRel AND #sSst AND #iPartPlaceOver_IFGantry;
END_REGION

REGION Network 30: STATE Num:60 Wait For Part Place By Gantry
   RUNG wire#powerrail
      Contact( #s60_WtPartPlaceByGantry )
      wire#w1
      I_Contact( #sStWtResetRel )
      I_Contact( #s60_WtPartPlaceByGantry_T1 )
      wire#w2
      Coil( #s60_WtPartPlaceByGantry )
   END_RUNG
   RUNG wire#powerrail
      Contact( #s50_WtShuttleRdyRcvPart_T1 )
   END_RUNG wire#w1
   RUNG wire#w2
      { S7_GenerateENO := "TRUE" } Move(in := 60, out1 => #StateNo)
   END_RUNG
   // the same network as SCL:
   #s60_WtPartPlaceByGantry := (#s60_WtPartPlaceByGantry OR #s50_WtShuttleRdyRcvPart_T1) AND NOT #sStWtResetRel AND NOT #s60_WtPartPlaceByGantry_T1;
   IF #s60_WtPartPlaceByGantry THEN #StateNo := 60; END_IF;
END_REGION

REGION Network 31: Actions for STATE Num:60 Wait For Part Place By Gantry
   RUNG wire#powerrail
      Contact( #s60_WtPartPlaceByGantry )
      Coil( #qInfeedGantry_PlaceStart )
   END_RUNG
   // the same network as SCL:
   #qInfeedGantry_PlaceStart := #s60_WtPartPlaceByGantry;
END_REGION

REGION Network 32: Condition1 for STATE Num:70 Check Part Present Status At Shuttle-1
   RUNG wire#powerrail
      I_Contact( #iPartPresent_Shuttle_1 )
      Coil( #c70_ChkPartPrsntStsShuttle1_T1 )
   END_RUNG
   // the same network as SCL:
   #c70_ChkPartPrsntStsShuttle1_T1 := NOT #iPartPresent_Shuttle_1;
END_REGION

REGION Network 33: Condition2 for STATE Num:70 Check Part Present Status At Shuttle-1
   RUNG wire#powerrail
      Contact( #iPartPresent_Shuttle_1 )
      Coil( #c70_ChkPartPrsntStsShuttle1_T2 )
   END_RUNG
   // the same network as SCL:
   #c70_ChkPartPrsntStsShuttle1_T2 := #iPartPresent_Shuttle_1;
END_REGION

REGION Network 34: Transition for STATE Num:70 Check Part Present Status At Shuttle-1
   RUNG wire#powerrail
      Contact( #s70_ChkPartPrsntStsShuttle1 )
      I_Contact( #sStWtResetRel )
      Contact( #sSst )
      wire#w1
      Contact( #c70_ChkPartPrsntStsShuttle1_T1 )
      Coil( #s70_ChkPartPrsntStsShuttle1_T1 )
   END_RUNG
   RUNG wire#w1
      I_Contact( #s70_ChkPartPrsntStsShuttle1_T1 )
      Contact( #c70_ChkPartPrsntStsShuttle1_T2 )
      Coil( #s70_ChkPartPrsntStsShuttle1_T2 )
   END_RUNG
   // the same network as SCL:
   #_w1 := #s70_ChkPartPrsntStsShuttle1 AND NOT #sStWtResetRel AND #sSst;
   #s70_ChkPartPrsntStsShuttle1_T1 := #_w1 AND #c70_ChkPartPrsntStsShuttle1_T1;
   #s70_ChkPartPrsntStsShuttle1_T2 := #_w1 AND NOT #s70_ChkPartPrsntStsShuttle1_T1 AND #c70_ChkPartPrsntStsShuttle1_T2;
END_REGION

REGION Network 35: STATE Num:70 Check Part Present Status At Shuttle-1
   RUNG wire#powerrail
      Contact( #s70_ChkPartPrsntStsShuttle1 )
      wire#w1
      I_Contact( #sStWtResetRel )
      I_Contact( #s70_ChkPartPrsntStsShuttle1_T1 )
      I_Contact( #s70_ChkPartPrsntStsShuttle1_T2 )
      wire#w2
      Coil( #s70_ChkPartPrsntStsShuttle1 )
   END_RUNG
   RUNG wire#powerrail
      Contact( #s120_WtPartUnldOvrTxGantry1_T1 )
   END_RUNG wire#w1
   RUNG wire#powerrail
      Contact( #s10_ChkPartStsAtSubStn_T3 )
   END_RUNG wire#w1
   RUNG wire#powerrail
      Contact( #s80_WtIFGantryPlacePart_T1 )
   END_RUNG wire#w1
   RUNG wire#w2
      { S7_GenerateENO := "TRUE" } Move(in := 70, out1 => #StateNo)
   END_RUNG
   // the same network as SCL:
   #s70_ChkPartPrsntStsShuttle1 := (#s70_ChkPartPrsntStsShuttle1 OR #s120_WtPartUnldOvrTxGantry1_T1 OR #s10_ChkPartStsAtSubStn_T3 OR #s80_WtIFGantryPlacePart_T1) AND NOT #sStWtResetRel AND NOT #s70_ChkPartPrsntStsShuttle1_T1 AND NOT #s70_ChkPartPrsntStsShuttle1_T2;
   IF #s70_ChkPartPrsntStsShuttle1 THEN #StateNo := 70; END_IF;
END_REGION

REGION Network 36: Transition for STATE Num:80 Wait for Infeed Gantry Place Part
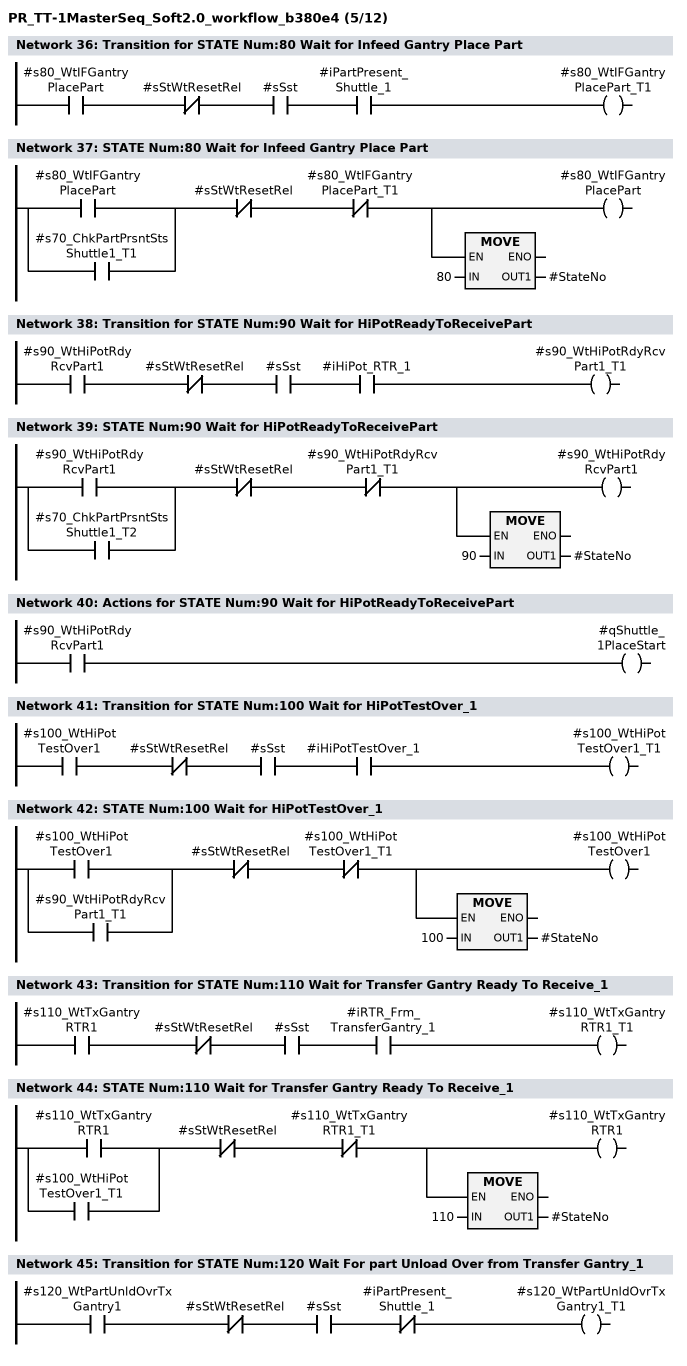
   RUNG wire#powerrail
      Contact( #s80_WtIFGantryPlacePart )
      I_Contact( #sStWtResetRel )
      Contact( #sSst )
      Contact( #iPartPresent_Shuttle_1 )
      Coil( #s80_WtIFGantryPlacePart_T1 )
   END_RUNG
   // the same network as SCL:
   #s80_WtIFGantryPlacePart_T1 := #s80_WtIFGantryPlacePart AND NOT #sStWtResetRel AND #sSst AND #iPartPresent_Shuttle_1;
END_REGION

REGION Network 37: STATE Num:80 Wait for Infeed Gantry Place Part
   RUNG wire#powerrail
      Contact( #s80_WtIFGantryPlacePart )
      wire#w1
      I_Contact( #sStWtResetRel )
      I_Contact( #s80_WtIFGantryPlacePart_T1 )
      wire#w2
      Coil( #s80_WtIFGantryPlacePart )
   END_RUNG
   RUNG wire#powerrail
      Contact( #s70_ChkPartPrsntStsShuttle1_T1 )
   END_RUNG wire#w1
   RUNG wire#w2
      { S7_GenerateENO := "TRUE" } Move(in := 80, out1 => #StateNo)
   END_RUNG
   // the same network as SCL:
   #s80_WtIFGantryPlacePart := (#s80_WtIFGantryPlacePart OR #s70_ChkPartPrsntStsShuttle1_T1) AND NOT #sStWtResetRel AND NOT #s80_WtIFGantryPlacePart_T1;
   IF #s80_WtIFGantryPlacePart THEN #StateNo := 80; END_IF;
END_REGION

REGION Network 38: Transition for STATE Num:90 Wait for HiPotReadyToReceivePart
   RUNG wire#powerrail
      Contact( #s90_WtHiPotRdyRcvPart1 )
      I_Contact( #sStWtResetRel )
      Contact( #sSst )
      Contact( #iHiPot_RTR_1 )
      Coil( #s90_WtHiPotRdyRcvPart1_T1 )
   END_RUNG
   // the same network as SCL:
   #s90_WtHiPotRdyRcvPart1_T1 := #s90_WtHiPotRdyRcvPart1 AND NOT #sStWtResetRel AND #sSst AND #iHiPot_RTR_1;
END_REGION

REGION Network 39: STATE Num:90 Wait for HiPotReadyToReceivePart
   RUNG wire#powerrail
      Contact( #s90_WtHiPotRdyRcvPart1 )
      wire#w1
      I_Contact( #sStWtResetRel )
      I_Contact( #s90_WtHiPotRdyRcvPart1_T1 )
      wire#w2
      Coil( #s90_WtHiPotRdyRcvPart1 )
   END_RUNG
   RUNG wire#powerrail
      Contact( #s70_ChkPartPrsntStsShuttle1_T2 )
   END_RUNG wire#w1
   RUNG wire#w2
      { S7_GenerateENO := "TRUE" } Move(in := 90, out1 => #StateNo)
   END_RUNG
   // the same network as SCL:
   #s90_WtHiPotRdyRcvPart1 := (#s90_WtHiPotRdyRcvPart1 OR #s70_ChkPartPrsntStsShuttle1_T2) AND NOT #sStWtResetRel AND NOT #s90_WtHiPotRdyRcvPart1_T1;
   IF #s90_WtHiPotRdyRcvPart1 THEN #StateNo := 90; END_IF;
END_REGION

REGION Network 40: Actions for STATE Num:90 Wait for HiPotReadyToReceivePart
   RUNG wire#powerrail
      Contact( #s90_WtHiPotRdyRcvPart1 )
      Coil( #qShuttle_1PlaceStart )
   END_RUNG
   // the same network as SCL:
   #qShuttle_1PlaceStart := #s90_WtHiPotRdyRcvPart1;
END_REGION

REGION Network 41: Transition for STATE Num:100 Wait for HiPotTestOver_1
   RUNG wire#powerrail
      Contact( #s100_WtHiPotTestOver1 )
      I_Contact( #sStWtResetRel )
      Contact( #sSst )
      Contact( #iHiPotTestOver_1 )
      Coil( #s100_WtHiPotTestOver1_T1 )
   END_RUNG
   // the same network as SCL:
   #s100_WtHiPotTestOver1_T1 := #s100_WtHiPotTestOver1 AND NOT #sStWtResetRel AND #sSst AND #iHiPotTestOver_1;
END_REGION

REGION Network 42: STATE Num:100 Wait for HiPotTestOver_1
   RUNG wire#powerrail
      Contact( #s100_WtHiPotTestOver1 )
      wire#w1
      I_Contact( #sStWtResetRel )
      I_Contact( #s100_WtHiPotTestOver1_T1 )
      wire#w2
      Coil( #s100_WtHiPotTestOver1 )
   END_RUNG
   RUNG wire#powerrail
      Contact( #s90_WtHiPotRdyRcvPart1_T1 )
   END_RUNG wire#w1
   RUNG wire#w2
      { S7_GenerateENO := "TRUE" } Move(in := 100, out1 => #StateNo)
   END_RUNG
   // the same network as SCL:
   #s100_WtHiPotTestOver1 := (#s100_WtHiPotTestOver1 OR #s90_WtHiPotRdyRcvPart1_T1) AND NOT #sStWtResetRel AND NOT #s100_WtHiPotTestOver1_T1;
   IF #s100_WtHiPotTestOver1 THEN #StateNo := 100; END_IF;
END_REGION

REGION Network 43: Transition for STATE Num:110 Wait for Transfer Gantry Ready To Receive_1
   RUNG wire#powerrail
      Contact( #s110_WtTxGantryRTR1 )
      I_Contact( #sStWtResetRel )
      Contact( #sSst )
      Contact( #iRTR_Frm_TransferGantry_1 )
      Coil( #s110_WtTxGantryRTR1_T1 )
   END_RUNG
   // the same network as SCL:
   #s110_WtTxGantryRTR1_T1 := #s110_WtTxGantryRTR1 AND NOT #sStWtResetRel AND #sSst AND #iRTR_Frm_TransferGantry_1;
END_REGION

REGION Network 44: STATE Num:110 Wait for Transfer Gantry Ready To Receive_1
   RUNG wire#powerrail
      Contact( #s110_WtTxGantryRTR1 )
      wire#w1
      I_Contact( #sStWtResetRel )
      I_Contact( #s110_WtTxGantryRTR1_T1 )
      wire#w2
      Coil( #s110_WtTxGantryRTR1 )
   END_RUNG
   RUNG wire#powerrail
      Contact( #s100_WtHiPotTestOver1_T1 )
   END_RUNG wire#w1
   RUNG wire#w2
      { S7_GenerateENO := "TRUE" } Move(in := 110, out1 => #StateNo)
   END_RUNG
   // the same network as SCL:
   #s110_WtTxGantryRTR1 := (#s110_WtTxGantryRTR1 OR #s100_WtHiPotTestOver1_T1) AND NOT #sStWtResetRel AND NOT #s110_WtTxGantryRTR1_T1;
   IF #s110_WtTxGantryRTR1 THEN #StateNo := 110; END_IF;
END_REGION

REGION Network 45: Transition for STATE Num:120 Wait For part Unload Over from Transfer Gantry_1
   RUNG wire#powerrail
      Contact( #s120_WtPartUnldOvrTxGantry1 )
      I_Contact( #sStWtResetRel )
      Contact( #sSst )
      I_Contact( #iPartPresent_Shuttle_1 )
      Coil( #s120_WtPartUnldOvrTxGantry1_T1 )
   END_RUNG
   // the same network as SCL:
   #s120_WtPartUnldOvrTxGantry1_T1 := #s120_WtPartUnldOvrTxGantry1 AND NOT #sStWtResetRel AND #sSst AND NOT #iPartPresent_Shuttle_1;
END_REGION

REGION Network 46: STATE Num:120 Wait For part Unload Over from Transfer Gantry_1
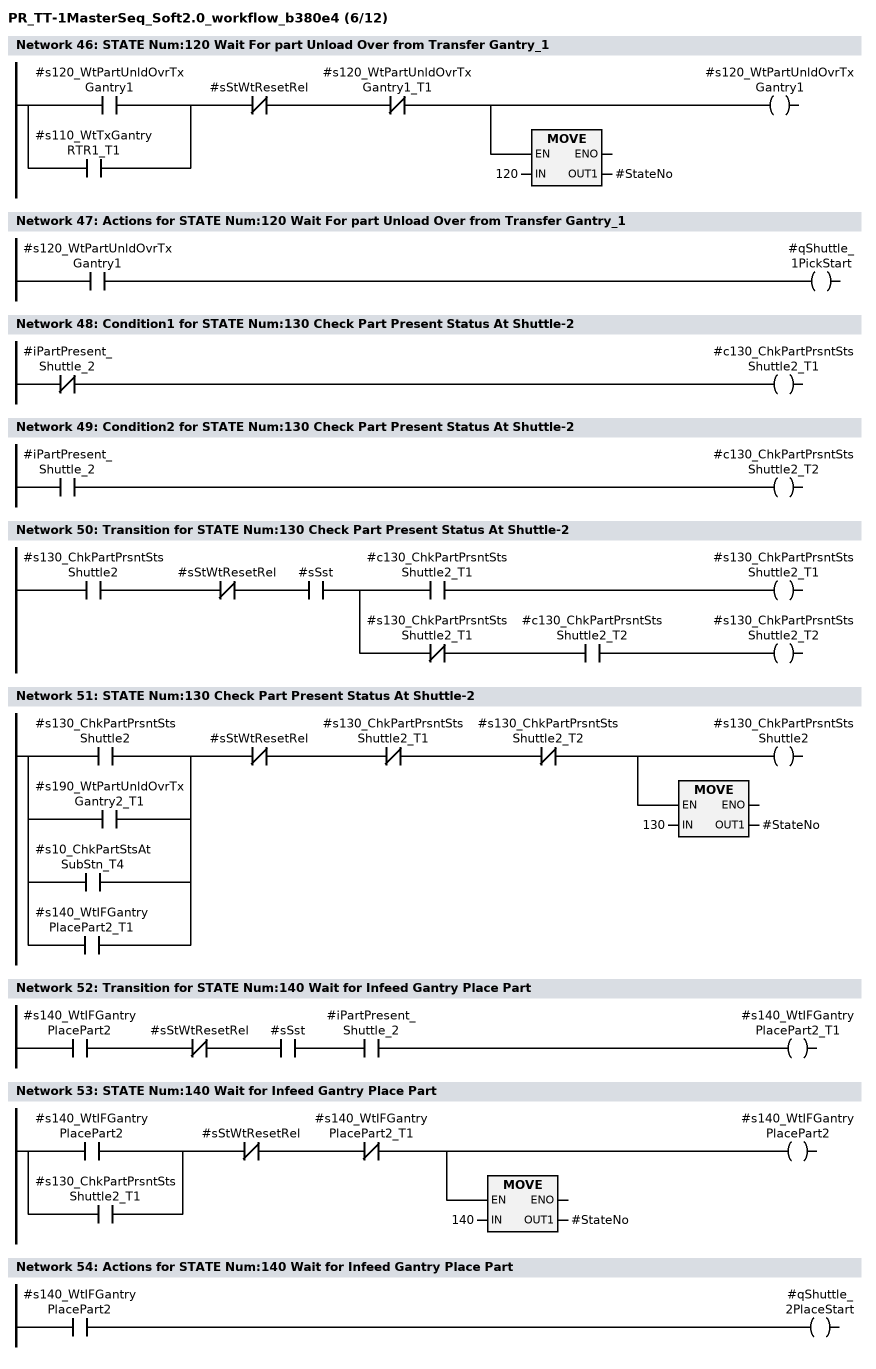
   RUNG wire#powerrail
      Contact( #s120_WtPartUnldOvrTxGantry1 )
      wire#w1
      I_Contact( #sStWtResetRel )
      I_Contact( #s120_WtPartUnldOvrTxGantry1_T1 )
      wire#w2
      Coil( #s120_WtPartUnldOvrTxGantry1 )
   END_RUNG
   RUNG wire#powerrail
      Contact( #s110_WtTxGantryRTR1_T1 )
   END_RUNG wire#w1
   RUNG wire#w2
      { S7_GenerateENO := "TRUE" } Move(in := 120, out1 => #StateNo)
   END_RUNG
   // the same network as SCL:
   #s120_WtPartUnldOvrTxGantry1 := (#s120_WtPartUnldOvrTxGantry1 OR #s110_WtTxGantryRTR1_T1) AND NOT #sStWtResetRel AND NOT #s120_WtPartUnldOvrTxGantry1_T1;
   IF #s120_WtPartUnldOvrTxGantry1 THEN #StateNo := 120; END_IF;
END_REGION

REGION Network 47: Actions for STATE Num:120 Wait For part Unload Over from Transfer Gantry_1
   RUNG wire#powerrail
      Contact( #s120_WtPartUnldOvrTxGantry1 )
      Coil( #qShuttle_1PickStart )
   END_RUNG
   // the same network as SCL:
   #qShuttle_1PickStart := #s120_WtPartUnldOvrTxGantry1;
END_REGION

REGION Network 48: Condition1 for STATE Num:130 Check Part Present Status At Shuttle-2
   RUNG wire#powerrail
      I_Contact( #iPartPresent_Shuttle_2 )
      Coil( #c130_ChkPartPrsntStsShuttle2_T1 )
   END_RUNG
   // the same network as SCL:
   #c130_ChkPartPrsntStsShuttle2_T1 := NOT #iPartPresent_Shuttle_2;
END_REGION

REGION Network 49: Condition2 for STATE Num:130 Check Part Present Status At Shuttle-2
   RUNG wire#powerrail
      Contact( #iPartPresent_Shuttle_2 )
      Coil( #c130_ChkPartPrsntStsShuttle2_T2 )
   END_RUNG
   // the same network as SCL:
   #c130_ChkPartPrsntStsShuttle2_T2 := #iPartPresent_Shuttle_2;
END_REGION

REGION Network 50: Transition for STATE Num:130 Check Part Present Status At Shuttle-2
   RUNG wire#powerrail
      Contact( #s130_ChkPartPrsntStsShuttle2 )
      I_Contact( #sStWtResetRel )
      Contact( #sSst )
      wire#w1
      Contact( #c130_ChkPartPrsntStsShuttle2_T1 )
      Coil( #s130_ChkPartPrsntStsShuttle2_T1 )
   END_RUNG
   RUNG wire#w1
      I_Contact( #s130_ChkPartPrsntStsShuttle2_T1 )
      Contact( #c130_ChkPartPrsntStsShuttle2_T2 )
      Coil( #s130_ChkPartPrsntStsShuttle2_T2 )
   END_RUNG
   // the same network as SCL:
   #_w1 := #s130_ChkPartPrsntStsShuttle2 AND NOT #sStWtResetRel AND #sSst;
   #s130_ChkPartPrsntStsShuttle2_T1 := #_w1 AND #c130_ChkPartPrsntStsShuttle2_T1;
   #s130_ChkPartPrsntStsShuttle2_T2 := #_w1 AND NOT #s130_ChkPartPrsntStsShuttle2_T1 AND #c130_ChkPartPrsntStsShuttle2_T2;
END_REGION

REGION Network 51: STATE Num:130 Check Part Present Status At Shuttle-2
   RUNG wire#powerrail
      Contact( #s130_ChkPartPrsntStsShuttle2 )
      wire#w1
      I_Contact( #sStWtResetRel )
      I_Contact( #s130_ChkPartPrsntStsShuttle2_T1 )
      I_Contact( #s130_ChkPartPrsntStsShuttle2_T2 )
      wire#w2
      Coil( #s130_ChkPartPrsntStsShuttle2 )
   END_RUNG
   RUNG wire#powerrail
      Contact( #s190_WtPartUnldOvrTxGantry2_T1 )
   END_RUNG wire#w1
   RUNG wire#powerrail
      Contact( #s10_ChkPartStsAtSubStn_T4 )
   END_RUNG wire#w1
   RUNG wire#powerrail
      Contact( #s140_WtIFGantryPlacePart2_T1 )
   END_RUNG wire#w1
   RUNG wire#w2
      { S7_GenerateENO := "TRUE" } Move(in := 130, out1 => #StateNo)
   END_RUNG
   // the same network as SCL:
   #s130_ChkPartPrsntStsShuttle2 := (#s130_ChkPartPrsntStsShuttle2 OR #s190_WtPartUnldOvrTxGantry2_T1 OR #s10_ChkPartStsAtSubStn_T4 OR #s140_WtIFGantryPlacePart2_T1) AND NOT #sStWtResetRel AND NOT #s130_ChkPartPrsntStsShuttle2_T1 AND NOT #s130_ChkPartPrsntStsShuttle2_T2;
   IF #s130_ChkPartPrsntStsShuttle2 THEN #StateNo := 130; END_IF;
END_REGION

REGION Network 52: Transition for STATE Num:140 Wait for Infeed Gantry Place Part
   RUNG wire#powerrail
      Contact( #s140_WtIFGantryPlacePart2 )
      I_Contact( #sStWtResetRel )
      Contact( #sSst )
      Contact( #iPartPresent_Shuttle_2 )
      Coil( #s140_WtIFGantryPlacePart2_T1 )
   END_RUNG
   // the same network as SCL:
   #s140_WtIFGantryPlacePart2_T1 := #s140_WtIFGantryPlacePart2 AND NOT #sStWtResetRel AND #sSst AND #iPartPresent_Shuttle_2;
END_REGION

REGION Network 53: STATE Num:140 Wait for Infeed Gantry Place Part
   RUNG wire#powerrail
      Contact( #s140_WtIFGantryPlacePart2 )
      wire#w1
      I_Contact( #sStWtResetRel )
      I_Contact( #s140_WtIFGantryPlacePart2_T1 )
      wire#w2
      Coil( #s140_WtIFGantryPlacePart2 )
   END_RUNG
   RUNG wire#powerrail
      Contact( #s130_ChkPartPrsntStsShuttle2_T1 )
   END_RUNG wire#w1
   RUNG wire#w2
      { S7_GenerateENO := "TRUE" } Move(in := 140, out1 => #StateNo)
   END_RUNG
   // the same network as SCL:
   #s140_WtIFGantryPlacePart2 := (#s140_WtIFGantryPlacePart2 OR #s130_ChkPartPrsntStsShuttle2_T1) AND NOT #sStWtResetRel AND NOT #s140_WtIFGantryPlacePart2_T1;
   IF #s140_WtIFGantryPlacePart2 THEN #StateNo := 140; END_IF;
END_REGION

REGION Network 54: Actions for STATE Num:140 Wait for Infeed Gantry Place Part
   RUNG wire#powerrail
      Contact( #s140_WtIFGantryPlacePart2 )
      Coil( #qShuttle_2PlaceStart )
   END_RUNG
   // the same network as SCL:
   #qShuttle_2PlaceStart := #s140_WtIFGantryPlacePart2;
END_REGION

REGION Network 55: Transition for STATE Num:150 Wait for HiPotReadyToReceivePart
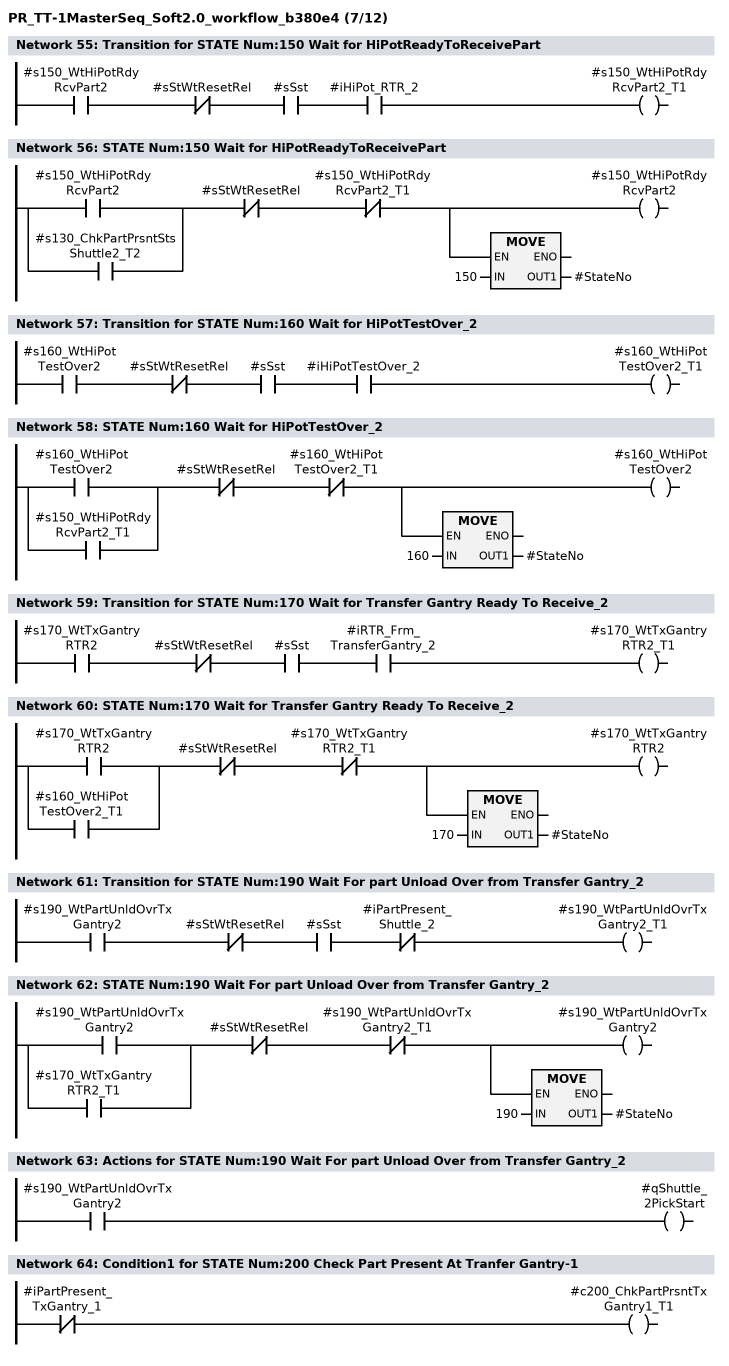
   RUNG wire#powerrail
      Contact( #s150_WtHiPotRdyRcvPart2 )
      I_Contact( #sStWtResetRel )
      Contact( #sSst )
      Contact( #iHiPot_RTR_2 )
      Coil( #s150_WtHiPotRdyRcvPart2_T1 )
   END_RUNG
   // the same network as SCL:
   #s150_WtHiPotRdyRcvPart2_T1 := #s150_WtHiPotRdyRcvPart2 AND NOT #sStWtResetRel AND #sSst AND #iHiPot_RTR_2;
END_REGION

REGION Network 56: STATE Num:150 Wait for HiPotReadyToReceivePart
   RUNG wire#powerrail
      Contact( #s150_WtHiPotRdyRcvPart2 )
      wire#w1
      I_Contact( #sStWtResetRel )
      I_Contact( #s150_WtHiPotRdyRcvPart2_T1 )
      wire#w2
      Coil( #s150_WtHiPotRdyRcvPart2 )
   END_RUNG
   RUNG wire#powerrail
      Contact( #s130_ChkPartPrsntStsShuttle2_T2 )
   END_RUNG wire#w1
   RUNG wire#w2
      { S7_GenerateENO := "TRUE" } Move(in := 150, out1 => #StateNo)
   END_RUNG
   // the same network as SCL:
   #s150_WtHiPotRdyRcvPart2 := (#s150_WtHiPotRdyRcvPart2 OR #s130_ChkPartPrsntStsShuttle2_T2) AND NOT #sStWtResetRel AND NOT #s150_WtHiPotRdyRcvPart2_T1;
   IF #s150_WtHiPotRdyRcvPart2 THEN #StateNo := 150; END_IF;
END_REGION

REGION Network 57: Transition for STATE Num:160 Wait for HiPotTestOver_2
   RUNG wire#powerrail
      Contact( #s160_WtHiPotTestOver2 )
      I_Contact( #sStWtResetRel )
      Contact( #sSst )
      Contact( #iHiPotTestOver_2 )
      Coil( #s160_WtHiPotTestOver2_T1 )
   END_RUNG
   // the same network as SCL:
   #s160_WtHiPotTestOver2_T1 := #s160_WtHiPotTestOver2 AND NOT #sStWtResetRel AND #sSst AND #iHiPotTestOver_2;
END_REGION

REGION Network 58: STATE Num:160 Wait for HiPotTestOver_2
   RUNG wire#powerrail
      Contact( #s160_WtHiPotTestOver2 )
      wire#w1
      I_Contact( #sStWtResetRel )
      I_Contact( #s160_WtHiPotTestOver2_T1 )
      wire#w2
      Coil( #s160_WtHiPotTestOver2 )
   END_RUNG
   RUNG wire#powerrail
      Contact( #s150_WtHiPotRdyRcvPart2_T1 )
   END_RUNG wire#w1
   RUNG wire#w2
      { S7_GenerateENO := "TRUE" } Move(in := 160, out1 => #StateNo)
   END_RUNG
   // the same network as SCL:
   #s160_WtHiPotTestOver2 := (#s160_WtHiPotTestOver2 OR #s150_WtHiPotRdyRcvPart2_T1) AND NOT #sStWtResetRel AND NOT #s160_WtHiPotTestOver2_T1;
   IF #s160_WtHiPotTestOver2 THEN #StateNo := 160; END_IF;
END_REGION

REGION Network 59: Transition for STATE Num:170 Wait for Transfer Gantry Ready To Receive_2
   RUNG wire#powerrail
      Contact( #s170_WtTxGantryRTR2 )
      I_Contact( #sStWtResetRel )
      Contact( #sSst )
      Contact( #iRTR_Frm_TransferGantry_2 )
      Coil( #s170_WtTxGantryRTR2_T1 )
   END_RUNG
   // the same network as SCL:
   #s170_WtTxGantryRTR2_T1 := #s170_WtTxGantryRTR2 AND NOT #sStWtResetRel AND #sSst AND #iRTR_Frm_TransferGantry_2;
END_REGION

REGION Network 60: STATE Num:170 Wait for Transfer Gantry Ready To Receive_2
   RUNG wire#powerrail
      Contact( #s170_WtTxGantryRTR2 )
      wire#w1
      I_Contact( #sStWtResetRel )
      I_Contact( #s170_WtTxGantryRTR2_T1 )
      wire#w2
      Coil( #s170_WtTxGantryRTR2 )
   END_RUNG
   RUNG wire#powerrail
      Contact( #s160_WtHiPotTestOver2_T1 )
   END_RUNG wire#w1
   RUNG wire#w2
      { S7_GenerateENO := "TRUE" } Move(in := 170, out1 => #StateNo)
   END_RUNG
   // the same network as SCL:
   #s170_WtTxGantryRTR2 := (#s170_WtTxGantryRTR2 OR #s160_WtHiPotTestOver2_T1) AND NOT #sStWtResetRel AND NOT #s170_WtTxGantryRTR2_T1;
   IF #s170_WtTxGantryRTR2 THEN #StateNo := 170; END_IF;
END_REGION

REGION Network 61: Transition for STATE Num:190 Wait For part Unload Over from Transfer Gantry_2
   RUNG wire#powerrail
      Contact( #s190_WtPartUnldOvrTxGantry2 )
      I_Contact( #sStWtResetRel )
      Contact( #sSst )
      I_Contact( #iPartPresent_Shuttle_2 )
      Coil( #s190_WtPartUnldOvrTxGantry2_T1 )
   END_RUNG
   // the same network as SCL:
   #s190_WtPartUnldOvrTxGantry2_T1 := #s190_WtPartUnldOvrTxGantry2 AND NOT #sStWtResetRel AND #sSst AND NOT #iPartPresent_Shuttle_2;
END_REGION

REGION Network 62: STATE Num:190 Wait For part Unload Over from Transfer Gantry_2
   RUNG wire#powerrail
      Contact( #s190_WtPartUnldOvrTxGantry2 )
      wire#w1
      I_Contact( #sStWtResetRel )
      I_Contact( #s190_WtPartUnldOvrTxGantry2_T1 )
      wire#w2
      Coil( #s190_WtPartUnldOvrTxGantry2 )
   END_RUNG
   RUNG wire#powerrail
      Contact( #s170_WtTxGantryRTR2_T1 )
   END_RUNG wire#w1
   RUNG wire#w2
      { S7_GenerateENO := "TRUE" } Move(in := 190, out1 => #StateNo)
   END_RUNG
   // the same network as SCL:
   #s190_WtPartUnldOvrTxGantry2 := (#s190_WtPartUnldOvrTxGantry2 OR #s170_WtTxGantryRTR2_T1) AND NOT #sStWtResetRel AND NOT #s190_WtPartUnldOvrTxGantry2_T1;
   IF #s190_WtPartUnldOvrTxGantry2 THEN #StateNo := 190; END_IF;
END_REGION

REGION Network 63: Actions for STATE Num:190 Wait For part Unload Over from Transfer Gantry_2
   RUNG wire#powerrail
      Contact( #s190_WtPartUnldOvrTxGantry2 )
      Coil( #qShuttle_2PickStart )
   END_RUNG
   // the same network as SCL:
   #qShuttle_2PickStart := #s190_WtPartUnldOvrTxGantry2;
END_REGION

REGION Network 64: Condition1 for STATE Num:200 Check Part Present At Tranfer Gantry-1
   RUNG wire#powerrail
      I_Contact( #iPartPresent_TxGantry_1 )
      Coil( #c200_ChkPartPrsntTxGantry1_T1 )
   END_RUNG
   // the same network as SCL:
   #c200_ChkPartPrsntTxGantry1_T1 := NOT #iPartPresent_TxGantry_1;
END_REGION

REGION Network 65: Condition2 for STATE Num:200 Check Part Present At Tranfer Gantry-1
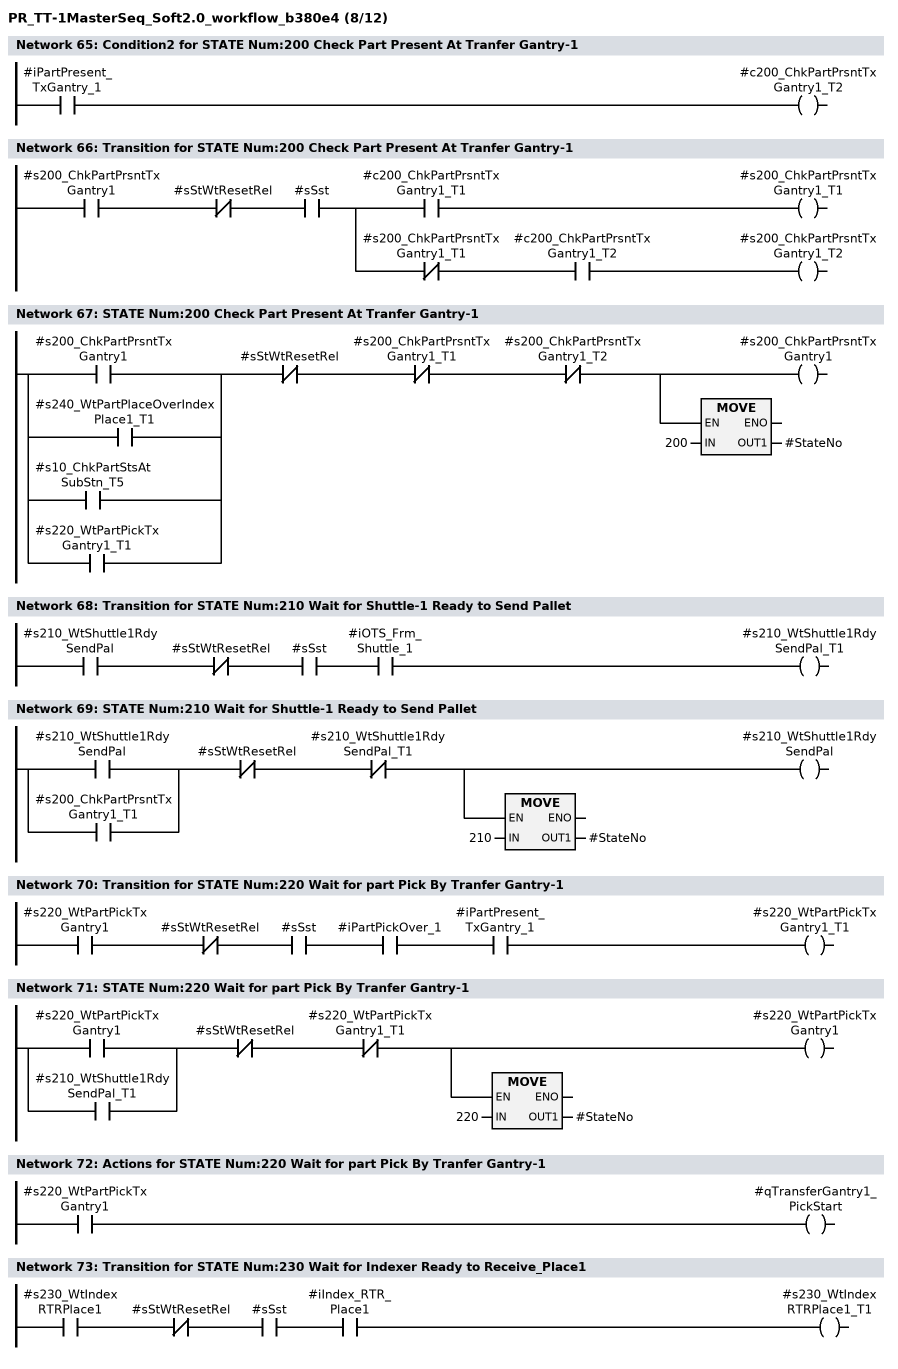
   RUNG wire#powerrail
      Contact( #iPartPresent_TxGantry_1 )
      Coil( #c200_ChkPartPrsntTxGantry1_T2 )
   END_RUNG
   // the same network as SCL:
   #c200_ChkPartPrsntTxGantry1_T2 := #iPartPresent_TxGantry_1;
END_REGION

REGION Network 66: Transition for STATE Num:200 Check Part Present At Tranfer Gantry-1
   RUNG wire#powerrail
      Contact( #s200_ChkPartPrsntTxGantry1 )
      I_Contact( #sStWtResetRel )
      Contact( #sSst )
      wire#w1
      Contact( #c200_ChkPartPrsntTxGantry1_T1 )
      Coil( #s200_ChkPartPrsntTxGantry1_T1 )
   END_RUNG
   RUNG wire#w1
      I_Contact( #s200_ChkPartPrsntTxGantry1_T1 )
      Contact( #c200_ChkPartPrsntTxGantry1_T2 )
      Coil( #s200_ChkPartPrsntTxGantry1_T2 )
   END_RUNG
   // the same network as SCL:
   #_w1 := #s200_ChkPartPrsntTxGantry1 AND NOT #sStWtResetRel AND #sSst;
   #s200_ChkPartPrsntTxGantry1_T1 := #_w1 AND #c200_ChkPartPrsntTxGantry1_T1;
   #s200_ChkPartPrsntTxGantry1_T2 := #_w1 AND NOT #s200_ChkPartPrsntTxGantry1_T1 AND #c200_ChkPartPrsntTxGantry1_T2;
END_REGION

REGION Network 67: STATE Num:200 Check Part Present At Tranfer Gantry-1
   RUNG wire#powerrail
      Contact( #s200_ChkPartPrsntTxGantry1 )
      wire#w1
      I_Contact( #sStWtResetRel )
      I_Contact( #s200_ChkPartPrsntTxGantry1_T1 )
      I_Contact( #s200_ChkPartPrsntTxGantry1_T2 )
      wire#w2
      Coil( #s200_ChkPartPrsntTxGantry1 )
   END_RUNG
   RUNG wire#powerrail
      Contact( #s240_WtPartPlaceOverIndexPlace1_T1 )
   END_RUNG wire#w1
   RUNG wire#powerrail
      Contact( #s10_ChkPartStsAtSubStn_T5 )
   END_RUNG wire#w1
   RUNG wire#powerrail
      Contact( #s220_WtPartPickTxGantry1_T1 )
   END_RUNG wire#w1
   RUNG wire#w2
      { S7_GenerateENO := "TRUE" } Move(in := 200, out1 => #StateNo)
   END_RUNG
   // the same network as SCL:
   #s200_ChkPartPrsntTxGantry1 := (#s200_ChkPartPrsntTxGantry1 OR #s240_WtPartPlaceOverIndexPlace1_T1 OR #s10_ChkPartStsAtSubStn_T5 OR #s220_WtPartPickTxGantry1_T1) AND NOT #sStWtResetRel AND NOT #s200_ChkPartPrsntTxGantry1_T1 AND NOT #s200_ChkPartPrsntTxGantry1_T2;
   IF #s200_ChkPartPrsntTxGantry1 THEN #StateNo := 200; END_IF;
END_REGION

REGION Network 68: Transition for STATE Num:210 Wait for Shuttle-1 Ready to Send Pallet
   RUNG wire#powerrail
      Contact( #s210_WtShuttle1RdySendPal )
      I_Contact( #sStWtResetRel )
      Contact( #sSst )
      Contact( #iOTS_Frm_Shuttle_1 )
      Coil( #s210_WtShuttle1RdySendPal_T1 )
   END_RUNG
   // the same network as SCL:
   #s210_WtShuttle1RdySendPal_T1 := #s210_WtShuttle1RdySendPal AND NOT #sStWtResetRel AND #sSst AND #iOTS_Frm_Shuttle_1;
END_REGION

REGION Network 69: STATE Num:210 Wait for Shuttle-1 Ready to Send Pallet
   RUNG wire#powerrail
      Contact( #s210_WtShuttle1RdySendPal )
      wire#w1
      I_Contact( #sStWtResetRel )
      I_Contact( #s210_WtShuttle1RdySendPal_T1 )
      wire#w2
      Coil( #s210_WtShuttle1RdySendPal )
   END_RUNG
   RUNG wire#powerrail
      Contact( #s200_ChkPartPrsntTxGantry1_T1 )
   END_RUNG wire#w1
   RUNG wire#w2
      { S7_GenerateENO := "TRUE" } Move(in := 210, out1 => #StateNo)
   END_RUNG
   // the same network as SCL:
   #s210_WtShuttle1RdySendPal := (#s210_WtShuttle1RdySendPal OR #s200_ChkPartPrsntTxGantry1_T1) AND NOT #sStWtResetRel AND NOT #s210_WtShuttle1RdySendPal_T1;
   IF #s210_WtShuttle1RdySendPal THEN #StateNo := 210; END_IF;
END_REGION

REGION Network 70: Transition for STATE Num:220 Wait for part Pick By Tranfer Gantry-1
   RUNG wire#powerrail
      Contact( #s220_WtPartPickTxGantry1 )
      I_Contact( #sStWtResetRel )
      Contact( #sSst )
      Contact( #iPartPickOver_1 )
      Contact( #iPartPresent_TxGantry_1 )
      Coil( #s220_WtPartPickTxGantry1_T1 )
   END_RUNG
   // the same network as SCL:
   #s220_WtPartPickTxGantry1_T1 := #s220_WtPartPickTxGantry1 AND NOT #sStWtResetRel AND #sSst AND #iPartPickOver_1 AND #iPartPresent_TxGantry_1;
END_REGION

REGION Network 71: STATE Num:220 Wait for part Pick By Tranfer Gantry-1
   RUNG wire#powerrail
      Contact( #s220_WtPartPickTxGantry1 )
      wire#w1
      I_Contact( #sStWtResetRel )
      I_Contact( #s220_WtPartPickTxGantry1_T1 )
      wire#w2
      Coil( #s220_WtPartPickTxGantry1 )
   END_RUNG
   RUNG wire#powerrail
      Contact( #s210_WtShuttle1RdySendPal_T1 )
   END_RUNG wire#w1
   RUNG wire#w2
      { S7_GenerateENO := "TRUE" } Move(in := 220, out1 => #StateNo)
   END_RUNG
   // the same network as SCL:
   #s220_WtPartPickTxGantry1 := (#s220_WtPartPickTxGantry1 OR #s210_WtShuttle1RdySendPal_T1) AND NOT #sStWtResetRel AND NOT #s220_WtPartPickTxGantry1_T1;
   IF #s220_WtPartPickTxGantry1 THEN #StateNo := 220; END_IF;
END_REGION

REGION Network 72: Actions for STATE Num:220 Wait for part Pick By Tranfer Gantry-1
   RUNG wire#powerrail
      Contact( #s220_WtPartPickTxGantry1 )
      Coil( #qTransferGantry1_PickStart )
   END_RUNG
   // the same network as SCL:
   #qTransferGantry1_PickStart := #s220_WtPartPickTxGantry1;
END_REGION

REGION Network 73: Transition for STATE Num:230 Wait for Indexer Ready to Receive_Place1
   RUNG wire#powerrail
      Contact( #s230_WtIndexRTRPlace1 )
      I_Contact( #sStWtResetRel )
      Contact( #sSst )
      Contact( #iIndex_RTR_Place1 )
      Coil( #s230_WtIndexRTRPlace1_T1 )
   END_RUNG
   // the same network as SCL:
   #s230_WtIndexRTRPlace1_T1 := #s230_WtIndexRTRPlace1 AND NOT #sStWtResetRel AND #sSst AND #iIndex_RTR_Place1;
END_REGION

REGION Network 74: STATE Num:230 Wait for Indexer Ready to Receive_Place1
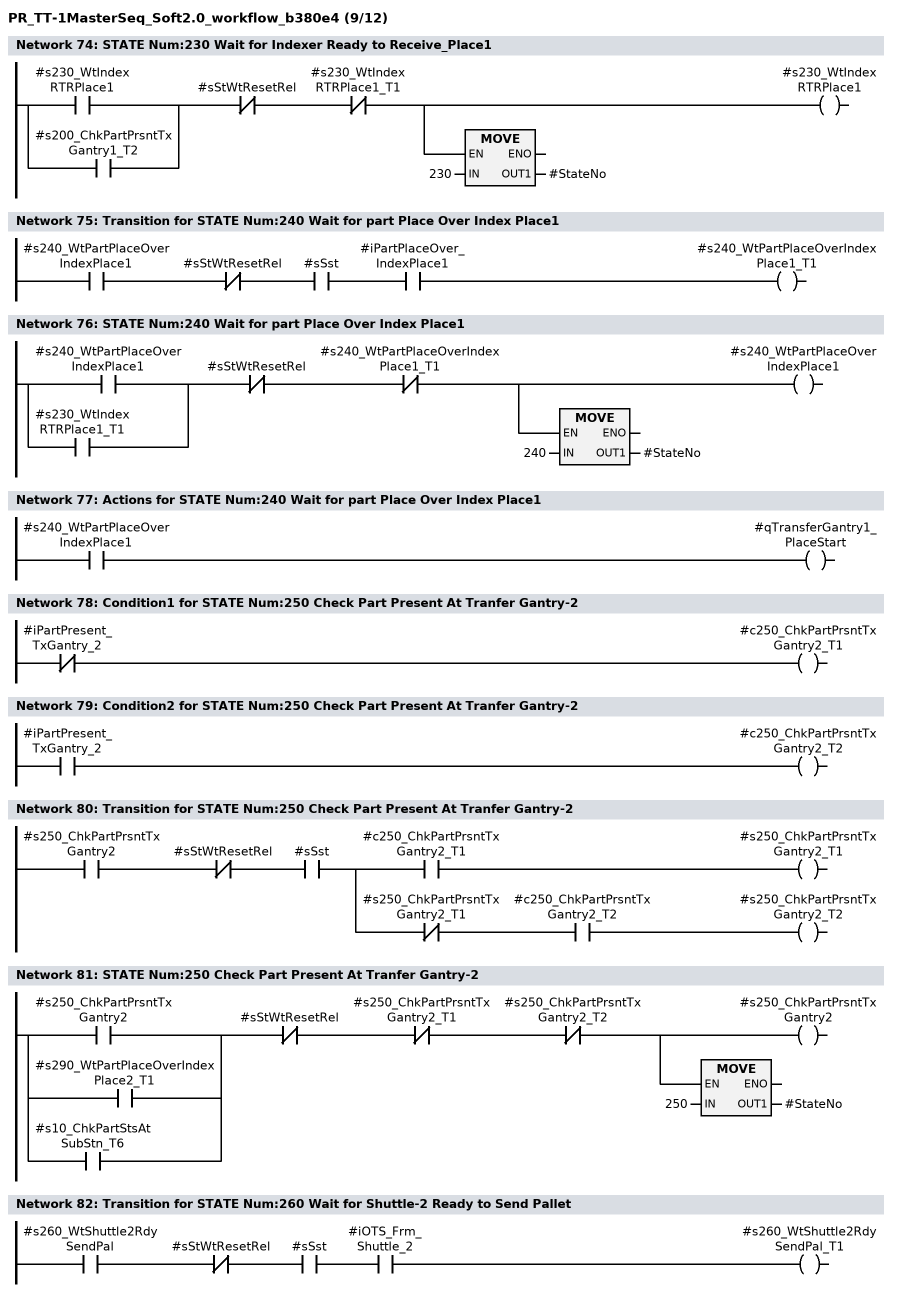
   RUNG wire#powerrail
      Contact( #s230_WtIndexRTRPlace1 )
      wire#w1
      I_Contact( #sStWtResetRel )
      I_Contact( #s230_WtIndexRTRPlace1_T1 )
      wire#w2
      Coil( #s230_WtIndexRTRPlace1 )
   END_RUNG
   RUNG wire#powerrail
      Contact( #s200_ChkPartPrsntTxGantry1_T2 )
   END_RUNG wire#w1
   RUNG wire#w2
      { S7_GenerateENO := "TRUE" } Move(in := 230, out1 => #StateNo)
   END_RUNG
   // the same network as SCL:
   #s230_WtIndexRTRPlace1 := (#s230_WtIndexRTRPlace1 OR #s200_ChkPartPrsntTxGantry1_T2) AND NOT #sStWtResetRel AND NOT #s230_WtIndexRTRPlace1_T1;
   IF #s230_WtIndexRTRPlace1 THEN #StateNo := 230; END_IF;
END_REGION

REGION Network 75: Transition for STATE Num:240 Wait for part Place Over Index Place1
   RUNG wire#powerrail
      Contact( #s240_WtPartPlaceOverIndexPlace1 )
      I_Contact( #sStWtResetRel )
      Contact( #sSst )
      Contact( #iPartPlaceOver_IndexPlace1 )
      Coil( #s240_WtPartPlaceOverIndexPlace1_T1 )
   END_RUNG
   // the same network as SCL:
   #s240_WtPartPlaceOverIndexPlace1_T1 := #s240_WtPartPlaceOverIndexPlace1 AND NOT #sStWtResetRel AND #sSst AND #iPartPlaceOver_IndexPlace1;
END_REGION

REGION Network 76: STATE Num:240 Wait for part Place Over Index Place1
   RUNG wire#powerrail
      Contact( #s240_WtPartPlaceOverIndexPlace1 )
      wire#w1
      I_Contact( #sStWtResetRel )
      I_Contact( #s240_WtPartPlaceOverIndexPlace1_T1 )
      wire#w2
      Coil( #s240_WtPartPlaceOverIndexPlace1 )
   END_RUNG
   RUNG wire#powerrail
      Contact( #s230_WtIndexRTRPlace1_T1 )
   END_RUNG wire#w1
   RUNG wire#w2
      { S7_GenerateENO := "TRUE" } Move(in := 240, out1 => #StateNo)
   END_RUNG
   // the same network as SCL:
   #s240_WtPartPlaceOverIndexPlace1 := (#s240_WtPartPlaceOverIndexPlace1 OR #s230_WtIndexRTRPlace1_T1) AND NOT #sStWtResetRel AND NOT #s240_WtPartPlaceOverIndexPlace1_T1;
   IF #s240_WtPartPlaceOverIndexPlace1 THEN #StateNo := 240; END_IF;
END_REGION

REGION Network 77: Actions for STATE Num:240 Wait for part Place Over Index Place1
   RUNG wire#powerrail
      Contact( #s240_WtPartPlaceOverIndexPlace1 )
      Coil( #qTransferGantry1_PlaceStart )
   END_RUNG
   // the same network as SCL:
   #qTransferGantry1_PlaceStart := #s240_WtPartPlaceOverIndexPlace1;
END_REGION

REGION Network 78: Condition1 for STATE Num:250 Check Part Present At Tranfer Gantry-2
   RUNG wire#powerrail
      I_Contact( #iPartPresent_TxGantry_2 )
      Coil( #c250_ChkPartPrsntTxGantry2_T1 )
   END_RUNG
   // the same network as SCL:
   #c250_ChkPartPrsntTxGantry2_T1 := NOT #iPartPresent_TxGantry_2;
END_REGION

REGION Network 79: Condition2 for STATE Num:250 Check Part Present At Tranfer Gantry-2
   RUNG wire#powerrail
      Contact( #iPartPresent_TxGantry_2 )
      Coil( #c250_ChkPartPrsntTxGantry2_T2 )
   END_RUNG
   // the same network as SCL:
   #c250_ChkPartPrsntTxGantry2_T2 := #iPartPresent_TxGantry_2;
END_REGION

REGION Network 80: Transition for STATE Num:250 Check Part Present At Tranfer Gantry-2
   RUNG wire#powerrail
      Contact( #s250_ChkPartPrsntTxGantry2 )
      I_Contact( #sStWtResetRel )
      Contact( #sSst )
      wire#w1
      Contact( #c250_ChkPartPrsntTxGantry2_T1 )
      Coil( #s250_ChkPartPrsntTxGantry2_T1 )
   END_RUNG
   RUNG wire#w1
      I_Contact( #s250_ChkPartPrsntTxGantry2_T1 )
      Contact( #c250_ChkPartPrsntTxGantry2_T2 )
      Coil( #s250_ChkPartPrsntTxGantry2_T2 )
   END_RUNG
   // the same network as SCL:
   #_w1 := #s250_ChkPartPrsntTxGantry2 AND NOT #sStWtResetRel AND #sSst;
   #s250_ChkPartPrsntTxGantry2_T1 := #_w1 AND #c250_ChkPartPrsntTxGantry2_T1;
   #s250_ChkPartPrsntTxGantry2_T2 := #_w1 AND NOT #s250_ChkPartPrsntTxGantry2_T1 AND #c250_ChkPartPrsntTxGantry2_T2;
END_REGION

REGION Network 81: STATE Num:250 Check Part Present At Tranfer Gantry-2
   RUNG wire#powerrail
      Contact( #s250_ChkPartPrsntTxGantry2 )
      wire#w1
      I_Contact( #sStWtResetRel )
      I_Contact( #s250_ChkPartPrsntTxGantry2_T1 )
      I_Contact( #s250_ChkPartPrsntTxGantry2_T2 )
      wire#w2
      Coil( #s250_ChkPartPrsntTxGantry2 )
   END_RUNG
   RUNG wire#powerrail
      Contact( #s290_WtPartPlaceOverIndexPlace2_T1 )
   END_RUNG wire#w1
   RUNG wire#powerrail
      Contact( #s10_ChkPartStsAtSubStn_T6 )
   END_RUNG wire#w1
   RUNG wire#w2
      { S7_GenerateENO := "TRUE" } Move(in := 250, out1 => #StateNo)
   END_RUNG
   // the same network as SCL:
   #s250_ChkPartPrsntTxGantry2 := (#s250_ChkPartPrsntTxGantry2 OR #s290_WtPartPlaceOverIndexPlace2_T1 OR #s10_ChkPartStsAtSubStn_T6) AND NOT #sStWtResetRel AND NOT #s250_ChkPartPrsntTxGantry2_T1 AND NOT #s250_ChkPartPrsntTxGantry2_T2;
   IF #s250_ChkPartPrsntTxGantry2 THEN #StateNo := 250; END_IF;
END_REGION

REGION Network 82: Transition for STATE Num:260 Wait for Shuttle-2 Ready to Send Pallet
   RUNG wire#powerrail
      Contact( #s260_WtShuttle2RdySendPal )
      I_Contact( #sStWtResetRel )
      Contact( #sSst )
      Contact( #iOTS_Frm_Shuttle_2 )
      Coil( #s260_WtShuttle2RdySendPal_T1 )
   END_RUNG
   // the same network as SCL:
   #s260_WtShuttle2RdySendPal_T1 := #s260_WtShuttle2RdySendPal AND NOT #sStWtResetRel AND #sSst AND #iOTS_Frm_Shuttle_2;
END_REGION

REGION Network 83: STATE Num:260 Wait for Shuttle-2 Ready to Send Pallet
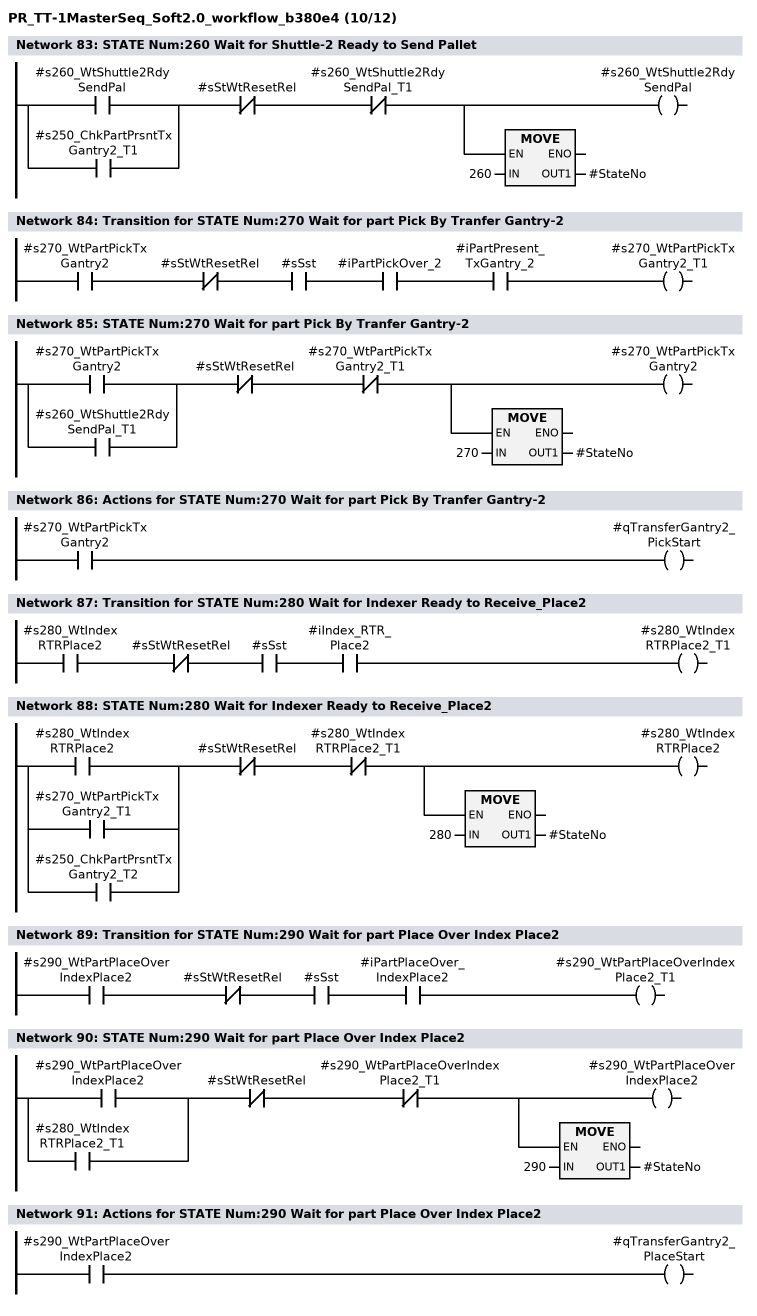
   RUNG wire#powerrail
      Contact( #s260_WtShuttle2RdySendPal )
      wire#w1
      I_Contact( #sStWtResetRel )
      I_Contact( #s260_WtShuttle2RdySendPal_T1 )
      wire#w2
      Coil( #s260_WtShuttle2RdySendPal )
   END_RUNG
   RUNG wire#powerrail
      Contact( #s250_ChkPartPrsntTxGantry2_T1 )
   END_RUNG wire#w1
   RUNG wire#w2
      { S7_GenerateENO := "TRUE" } Move(in := 260, out1 => #StateNo)
   END_RUNG
   // the same network as SCL:
   #s260_WtShuttle2RdySendPal := (#s260_WtShuttle2RdySendPal OR #s250_ChkPartPrsntTxGantry2_T1) AND NOT #sStWtResetRel AND NOT #s260_WtShuttle2RdySendPal_T1;
   IF #s260_WtShuttle2RdySendPal THEN #StateNo := 260; END_IF;
END_REGION

REGION Network 84: Transition for STATE Num:270 Wait for part Pick By Tranfer Gantry-2
   RUNG wire#powerrail
      Contact( #s270_WtPartPickTxGantry2 )
      I_Contact( #sStWtResetRel )
      Contact( #sSst )
      Contact( #iPartPickOver_2 )
      Contact( #iPartPresent_TxGantry_2 )
      Coil( #s270_WtPartPickTxGantry2_T1 )
   END_RUNG
   // the same network as SCL:
   #s270_WtPartPickTxGantry2_T1 := #s270_WtPartPickTxGantry2 AND NOT #sStWtResetRel AND #sSst AND #iPartPickOver_2 AND #iPartPresent_TxGantry_2;
END_REGION

REGION Network 85: STATE Num:270 Wait for part Pick By Tranfer Gantry-2
   RUNG wire#powerrail
      Contact( #s270_WtPartPickTxGantry2 )
      wire#w1
      I_Contact( #sStWtResetRel )
      I_Contact( #s270_WtPartPickTxGantry2_T1 )
      wire#w2
      Coil( #s270_WtPartPickTxGantry2 )
   END_RUNG
   RUNG wire#powerrail
      Contact( #s260_WtShuttle2RdySendPal_T1 )
   END_RUNG wire#w1
   RUNG wire#w2
      { S7_GenerateENO := "TRUE" } Move(in := 270, out1 => #StateNo)
   END_RUNG
   // the same network as SCL:
   #s270_WtPartPickTxGantry2 := (#s270_WtPartPickTxGantry2 OR #s260_WtShuttle2RdySendPal_T1) AND NOT #sStWtResetRel AND NOT #s270_WtPartPickTxGantry2_T1;
   IF #s270_WtPartPickTxGantry2 THEN #StateNo := 270; END_IF;
END_REGION

REGION Network 86: Actions for STATE Num:270 Wait for part Pick By Tranfer Gantry-2
   RUNG wire#powerrail
      Contact( #s270_WtPartPickTxGantry2 )
      Coil( #qTransferGantry2_PickStart )
   END_RUNG
   // the same network as SCL:
   #qTransferGantry2_PickStart := #s270_WtPartPickTxGantry2;
END_REGION

REGION Network 87: Transition for STATE Num:280 Wait for Indexer Ready to Receive_Place2
   RUNG wire#powerrail
      Contact( #s280_WtIndexRTRPlace2 )
      I_Contact( #sStWtResetRel )
      Contact( #sSst )
      Contact( #iIndex_RTR_Place2 )
      Coil( #s280_WtIndexRTRPlace2_T1 )
   END_RUNG
   // the same network as SCL:
   #s280_WtIndexRTRPlace2_T1 := #s280_WtIndexRTRPlace2 AND NOT #sStWtResetRel AND #sSst AND #iIndex_RTR_Place2;
END_REGION

REGION Network 88: STATE Num:280 Wait for Indexer Ready to Receive_Place2
   RUNG wire#powerrail
      Contact( #s280_WtIndexRTRPlace2 )
      wire#w1
      I_Contact( #sStWtResetRel )
      I_Contact( #s280_WtIndexRTRPlace2_T1 )
      wire#w2
      Coil( #s280_WtIndexRTRPlace2 )
   END_RUNG
   RUNG wire#powerrail
      Contact( #s270_WtPartPickTxGantry2_T1 )
   END_RUNG wire#w1
   RUNG wire#powerrail
      Contact( #s250_ChkPartPrsntTxGantry2_T2 )
   END_RUNG wire#w1
   RUNG wire#w2
      { S7_GenerateENO := "TRUE" } Move(in := 280, out1 => #StateNo)
   END_RUNG
   // the same network as SCL:
   #s280_WtIndexRTRPlace2 := (#s280_WtIndexRTRPlace2 OR #s270_WtPartPickTxGantry2_T1 OR #s250_ChkPartPrsntTxGantry2_T2) AND NOT #sStWtResetRel AND NOT #s280_WtIndexRTRPlace2_T1;
   IF #s280_WtIndexRTRPlace2 THEN #StateNo := 280; END_IF;
END_REGION

REGION Network 89: Transition for STATE Num:290 Wait for part Place Over Index Place2
   RUNG wire#powerrail
      Contact( #s290_WtPartPlaceOverIndexPlace2 )
      I_Contact( #sStWtResetRel )
      Contact( #sSst )
      Contact( #iPartPlaceOver_IndexPlace2 )
      Coil( #s290_WtPartPlaceOverIndexPlace2_T1 )
   END_RUNG
   // the same network as SCL:
   #s290_WtPartPlaceOverIndexPlace2_T1 := #s290_WtPartPlaceOverIndexPlace2 AND NOT #sStWtResetRel AND #sSst AND #iPartPlaceOver_IndexPlace2;
END_REGION

REGION Network 90: STATE Num:290 Wait for part Place Over Index Place2
   RUNG wire#powerrail
      Contact( #s290_WtPartPlaceOverIndexPlace2 )
      wire#w1
      I_Contact( #sStWtResetRel )
      I_Contact( #s290_WtPartPlaceOverIndexPlace2_T1 )
      wire#w2
      Coil( #s290_WtPartPlaceOverIndexPlace2 )
   END_RUNG
   RUNG wire#powerrail
      Contact( #s280_WtIndexRTRPlace2_T1 )
   END_RUNG wire#w1
   RUNG wire#w2
      { S7_GenerateENO := "TRUE" } Move(in := 290, out1 => #StateNo)
   END_RUNG
   // the same network as SCL:
   #s290_WtPartPlaceOverIndexPlace2 := (#s290_WtPartPlaceOverIndexPlace2 OR #s280_WtIndexRTRPlace2_T1) AND NOT #sStWtResetRel AND NOT #s290_WtPartPlaceOverIndexPlace2_T1;
   IF #s290_WtPartPlaceOverIndexPlace2 THEN #StateNo := 290; END_IF;
END_REGION

REGION Network 91: Actions for STATE Num:290 Wait for part Place Over Index Place2
   RUNG wire#powerrail
      Contact( #s290_WtPartPlaceOverIndexPlace2 )
      Coil( #qTransferGantry2_PlaceStart )
   END_RUNG
   // the same network as SCL:
   #qTransferGantry2_PlaceStart := #s290_WtPartPlaceOverIndexPlace2;
END_REGION

REGION Network 92: Condition1 for STATE Num:300 Check Part Present At Indexer
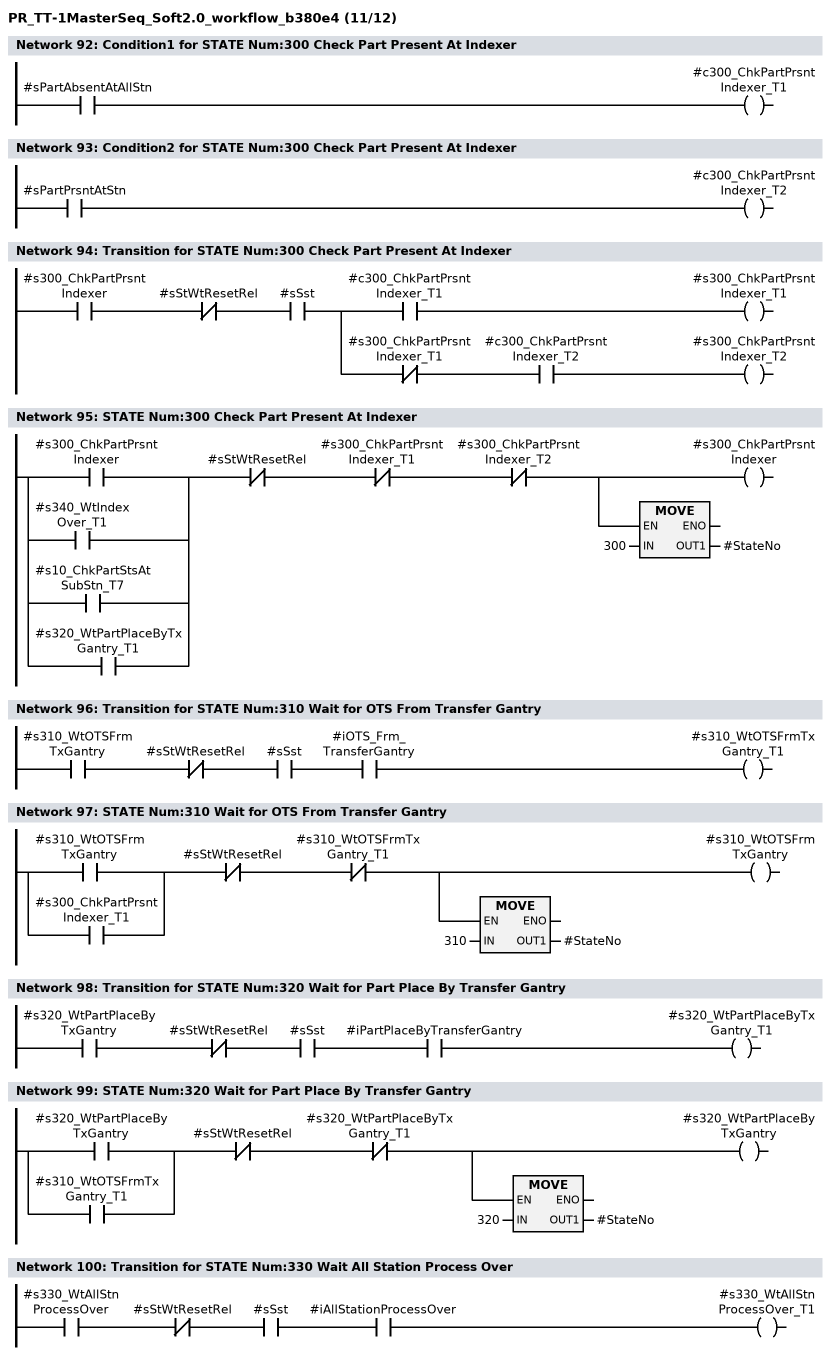
   RUNG wire#powerrail
      Contact( #sPartAbsentAtAllStn )
      Coil( #c300_ChkPartPrsntIndexer_T1 )
   END_RUNG
   // the same network as SCL:
   #c300_ChkPartPrsntIndexer_T1 := #sPartAbsentAtAllStn;
END_REGION

REGION Network 93: Condition2 for STATE Num:300 Check Part Present At Indexer
   RUNG wire#powerrail
      Contact( #sPartPrsntAtStn )
      Coil( #c300_ChkPartPrsntIndexer_T2 )
   END_RUNG
   // the same network as SCL:
   #c300_ChkPartPrsntIndexer_T2 := #sPartPrsntAtStn;
END_REGION

REGION Network 94: Transition for STATE Num:300 Check Part Present At Indexer
   RUNG wire#powerrail
      Contact( #s300_ChkPartPrsntIndexer )
      I_Contact( #sStWtResetRel )
      Contact( #sSst )
      wire#w1
      Contact( #c300_ChkPartPrsntIndexer_T1 )
      Coil( #s300_ChkPartPrsntIndexer_T1 )
   END_RUNG
   RUNG wire#w1
      I_Contact( #s300_ChkPartPrsntIndexer_T1 )
      Contact( #c300_ChkPartPrsntIndexer_T2 )
      Coil( #s300_ChkPartPrsntIndexer_T2 )
   END_RUNG
   // the same network as SCL:
   #_w1 := #s300_ChkPartPrsntIndexer AND NOT #sStWtResetRel AND #sSst;
   #s300_ChkPartPrsntIndexer_T1 := #_w1 AND #c300_ChkPartPrsntIndexer_T1;
   #s300_ChkPartPrsntIndexer_T2 := #_w1 AND NOT #s300_ChkPartPrsntIndexer_T1 AND #c300_ChkPartPrsntIndexer_T2;
END_REGION

REGION Network 95: STATE Num:300 Check Part Present At Indexer
   RUNG wire#powerrail
      Contact( #s300_ChkPartPrsntIndexer )
      wire#w1
      I_Contact( #sStWtResetRel )
      I_Contact( #s300_ChkPartPrsntIndexer_T1 )
      I_Contact( #s300_ChkPartPrsntIndexer_T2 )
      wire#w2
      Coil( #s300_ChkPartPrsntIndexer )
   END_RUNG
   RUNG wire#powerrail
      Contact( #s340_WtIndexOver_T1 )
   END_RUNG wire#w1
   RUNG wire#powerrail
      Contact( #s10_ChkPartStsAtSubStn_T7 )
   END_RUNG wire#w1
   RUNG wire#powerrail
      Contact( #s320_WtPartPlaceByTxGantry_T1 )
   END_RUNG wire#w1
   RUNG wire#w2
      { S7_GenerateENO := "TRUE" } Move(in := 300, out1 => #StateNo)
   END_RUNG
   // the same network as SCL:
   #s300_ChkPartPrsntIndexer := (#s300_ChkPartPrsntIndexer OR #s340_WtIndexOver_T1 OR #s10_ChkPartStsAtSubStn_T7 OR #s320_WtPartPlaceByTxGantry_T1) AND NOT #sStWtResetRel AND NOT #s300_ChkPartPrsntIndexer_T1 AND NOT #s300_ChkPartPrsntIndexer_T2;
   IF #s300_ChkPartPrsntIndexer THEN #StateNo := 300; END_IF;
END_REGION

REGION Network 96: Transition for STATE Num:310 Wait for OTS From Transfer Gantry
   RUNG wire#powerrail
      Contact( #s310_WtOTSFrmTxGantry )
      I_Contact( #sStWtResetRel )
      Contact( #sSst )
      Contact( #iOTS_Frm_TransferGantry )
      Coil( #s310_WtOTSFrmTxGantry_T1 )
   END_RUNG
   // the same network as SCL:
   #s310_WtOTSFrmTxGantry_T1 := #s310_WtOTSFrmTxGantry AND NOT #sStWtResetRel AND #sSst AND #iOTS_Frm_TransferGantry;
END_REGION

REGION Network 97: STATE Num:310 Wait for OTS From Transfer Gantry
   RUNG wire#powerrail
      Contact( #s310_WtOTSFrmTxGantry )
      wire#w1
      I_Contact( #sStWtResetRel )
      I_Contact( #s310_WtOTSFrmTxGantry_T1 )
      wire#w2
      Coil( #s310_WtOTSFrmTxGantry )
   END_RUNG
   RUNG wire#powerrail
      Contact( #s300_ChkPartPrsntIndexer_T1 )
   END_RUNG wire#w1
   RUNG wire#w2
      { S7_GenerateENO := "TRUE" } Move(in := 310, out1 => #StateNo)
   END_RUNG
   // the same network as SCL:
   #s310_WtOTSFrmTxGantry := (#s310_WtOTSFrmTxGantry OR #s300_ChkPartPrsntIndexer_T1) AND NOT #sStWtResetRel AND NOT #s310_WtOTSFrmTxGantry_T1;
   IF #s310_WtOTSFrmTxGantry THEN #StateNo := 310; END_IF;
END_REGION

REGION Network 98: Transition for STATE Num:320 Wait for Part Place By Transfer Gantry
   RUNG wire#powerrail
      Contact( #s320_WtPartPlaceByTxGantry )
      I_Contact( #sStWtResetRel )
      Contact( #sSst )
      Contact( #iPartPlaceByTransferGantry )
      Coil( #s320_WtPartPlaceByTxGantry_T1 )
   END_RUNG
   // the same network as SCL:
   #s320_WtPartPlaceByTxGantry_T1 := #s320_WtPartPlaceByTxGantry AND NOT #sStWtResetRel AND #sSst AND #iPartPlaceByTransferGantry;
END_REGION

REGION Network 99: STATE Num:320 Wait for Part Place By Transfer Gantry
   RUNG wire#powerrail
      Contact( #s320_WtPartPlaceByTxGantry )
      wire#w1
      I_Contact( #sStWtResetRel )
      I_Contact( #s320_WtPartPlaceByTxGantry_T1 )
      wire#w2
      Coil( #s320_WtPartPlaceByTxGantry )
   END_RUNG
   RUNG wire#powerrail
      Contact( #s310_WtOTSFrmTxGantry_T1 )
   END_RUNG wire#w1
   RUNG wire#w2
      { S7_GenerateENO := "TRUE" } Move(in := 320, out1 => #StateNo)
   END_RUNG
   // the same network as SCL:
   #s320_WtPartPlaceByTxGantry := (#s320_WtPartPlaceByTxGantry OR #s310_WtOTSFrmTxGantry_T1) AND NOT #sStWtResetRel AND NOT #s320_WtPartPlaceByTxGantry_T1;
   IF #s320_WtPartPlaceByTxGantry THEN #StateNo := 320; END_IF;
END_REGION

REGION Network 100: Transition for STATE Num:330 Wait All Station Process Over
   RUNG wire#powerrail
      Contact( #s330_WtAllStnProcessOver )
      I_Contact( #sStWtResetRel )
      Contact( #sSst )
      Contact( #iAllStationProcessOver )
      Coil( #s330_WtAllStnProcessOver_T1 )
   END_RUNG
   // the same network as SCL:
   #s330_WtAllStnProcessOver_T1 := #s330_WtAllStnProcessOver AND NOT #sStWtResetRel AND #sSst AND #iAllStationProcessOver;
END_REGION

REGION Network 101: STATE Num:330 Wait All Station Process Over
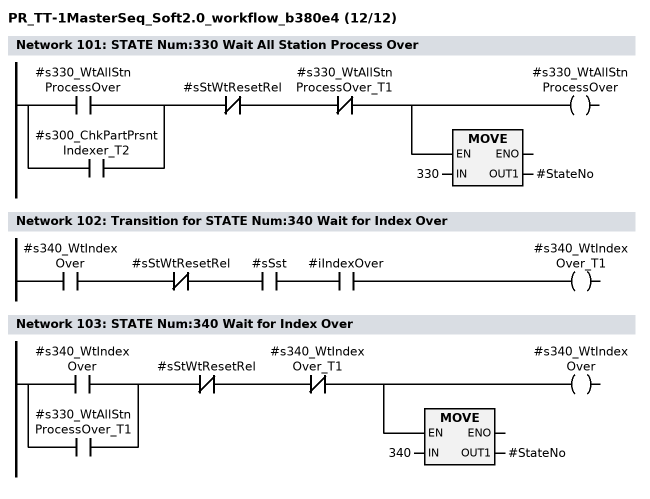
   RUNG wire#powerrail
      Contact( #s330_WtAllStnProcessOver )
      wire#w1
      I_Contact( #sStWtResetRel )
      I_Contact( #s330_WtAllStnProcessOver_T1 )
      wire#w2
      Coil( #s330_WtAllStnProcessOver )
   END_RUNG
   RUNG wire#powerrail
      Contact( #s300_ChkPartPrsntIndexer_T2 )
   END_RUNG wire#w1
   RUNG wire#w2
      { S7_GenerateENO := "TRUE" } Move(in := 330, out1 => #StateNo)
   END_RUNG
   // the same network as SCL:
   #s330_WtAllStnProcessOver := (#s330_WtAllStnProcessOver OR #s300_ChkPartPrsntIndexer_T2) AND NOT #sStWtResetRel AND NOT #s330_WtAllStnProcessOver_T1;
   IF #s330_WtAllStnProcessOver THEN #StateNo := 330; END_IF;
END_REGION

REGION Network 102: Transition for STATE Num:340 Wait for Index Over
   RUNG wire#powerrail
      Contact( #s340_WtIndexOver )
      I_Contact( #sStWtResetRel )
      Contact( #sSst )
      Contact( #iIndexOver )
      Coil( #s340_WtIndexOver_T1 )
   END_RUNG
   // the same network as SCL:
   #s340_WtIndexOver_T1 := #s340_WtIndexOver AND NOT #sStWtResetRel AND #sSst AND #iIndexOver;
END_REGION

REGION Network 103: STATE Num:340 Wait for Index Over
   RUNG wire#powerrail
      Contact( #s340_WtIndexOver )
      wire#w1
      I_Contact( #sStWtResetRel )
      I_Contact( #s340_WtIndexOver_T1 )
      wire#w2
      Coil( #s340_WtIndexOver )
   END_RUNG
   RUNG wire#powerrail
      Contact( #s330_WtAllStnProcessOver_T1 )
   END_RUNG wire#w1
   RUNG wire#w2
      { S7_GenerateENO := "TRUE" } Move(in := 340, out1 => #StateNo)
   END_RUNG
   // the same network as SCL:
   #s340_WtIndexOver := (#s340_WtIndexOver OR #s330_WtAllStnProcessOver_T1) AND NOT #sStWtResetRel AND NOT #s340_WtIndexOver_T1;
   IF #s340_WtIndexOver THEN #StateNo := 340; END_IF;
END_REGION
END_FUNCTION_BLOCK
